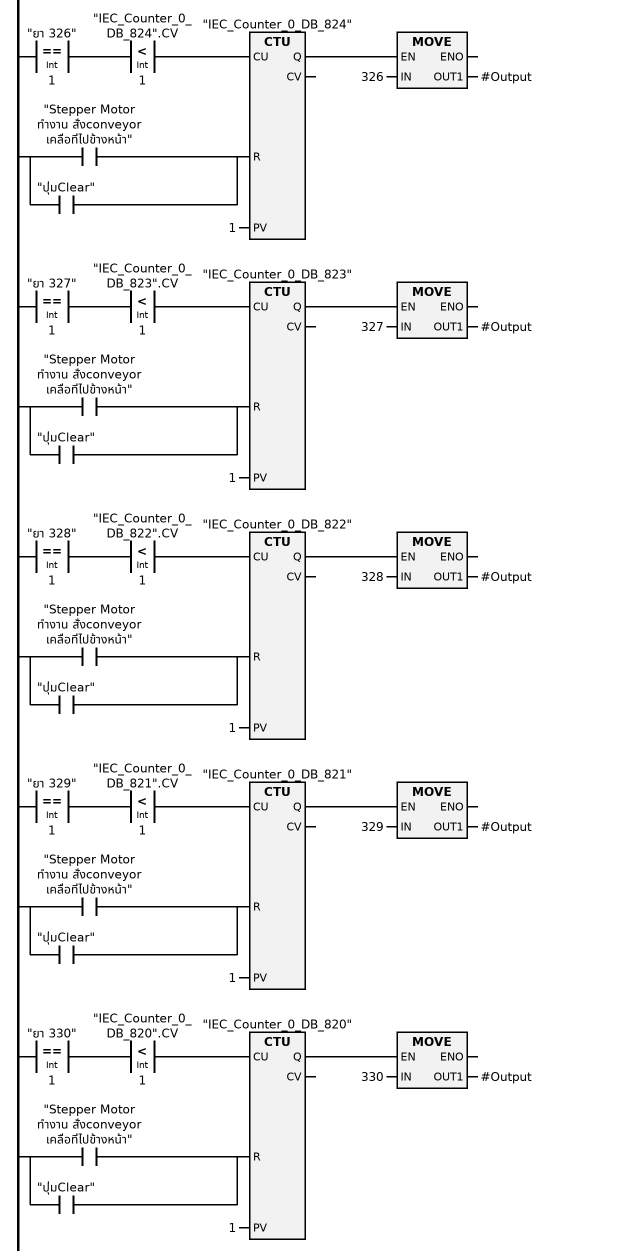
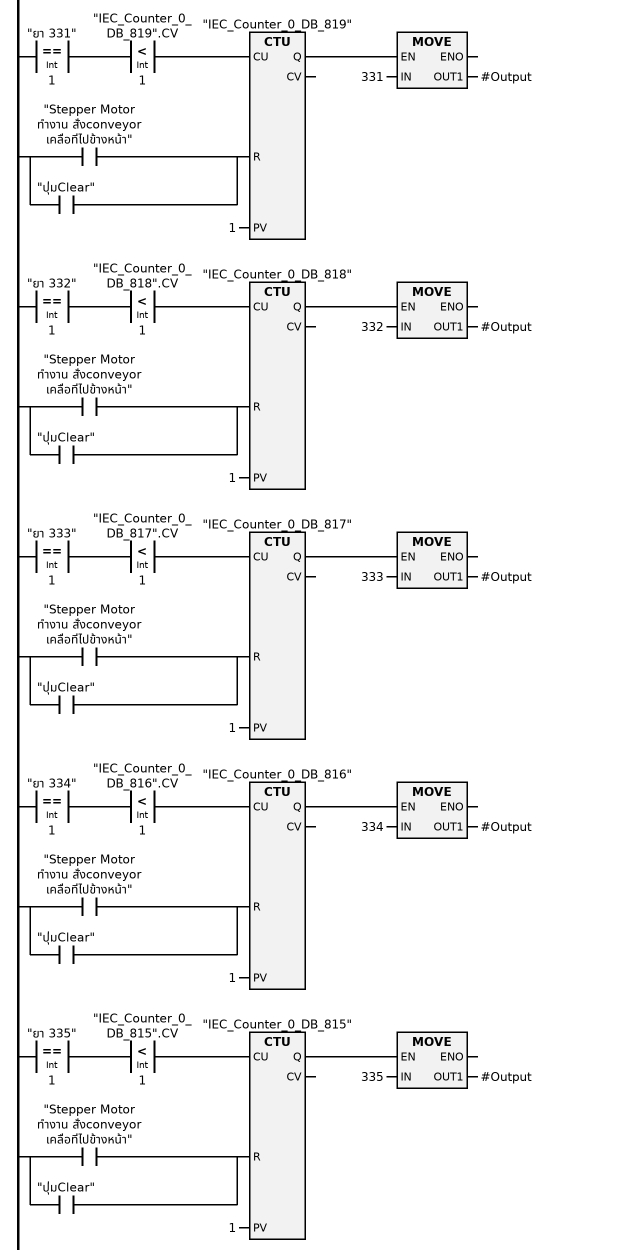
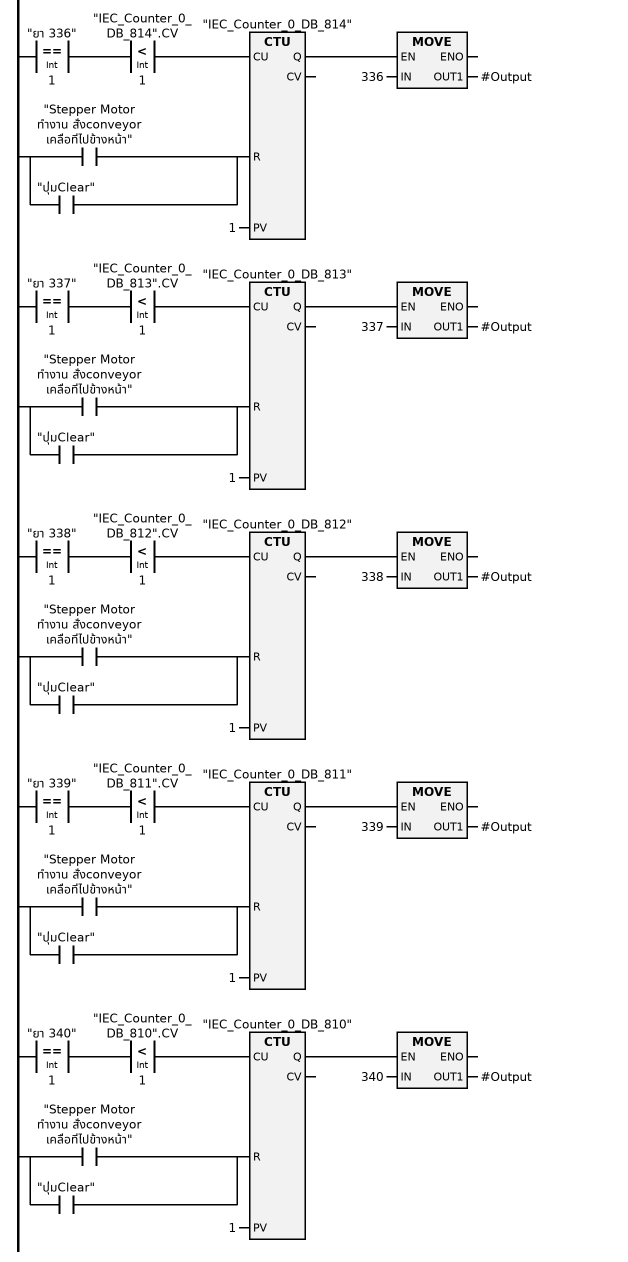
   "IEC_Counter_0_DB_829".CTU(CU := ("ยา 321" = 1) AND ("IEC_Counter_0_DB_829".CV < 1),
                           R := "Stepper Motor ทำงาน สั่งconveyor เคลื่อที่ไปข้างหน้า" OR "ปุ่มClear",
                           PV := 1);
   IF "IEC_Counter_0_DB_829".Q THEN #Output := 321; END_IF;
   "IEC_Counter_0_DB_828".CTU(CU := ("ยา 322" = 1) AND ("IEC_Counter_0_DB_828".CV < 1),
                           R := "Stepper Motor ทำงาน สั่งconveyor เคลื่อที่ไปข้างหน้า" OR "ปุ่มClear",
                           PV := 1);
   IF "IEC_Counter_0_DB_828".Q THEN #Output := 322; END_IF;
   "IEC_Counter_0_DB_825".CTU(CU := ("ยา 323" = 1) AND ("IEC_Counter_0_DB_825".CV < 1),
                           R := "Stepper Motor ทำงาน สั่งconveyor เคลื่อที่ไปข้างหน้า" OR "ปุ่มClear",
                           PV := 1);
   IF "IEC_Counter_0_DB_825".Q THEN #Output := 323; END_IF;
   "IEC_Counter_0_DB_827".CTU(CU := ("ยา 324" = 1) AND ("IEC_Counter_0_DB_827".CV < 1),
                           R := "Stepper Motor ทำงาน สั่งconveyor เคลื่อที่ไปข้างหน้า" OR "ปุ่มClear",
                           PV := 1);
   IF "IEC_Counter_0_DB_827".Q THEN #Output := 324; END_IF;
   "IEC_Counter_0_DB_826".CTU(CU := ("ยา 325" = 1) AND ("IEC_Counter_0_DB_826".CV < 1),
                           R := "Stepper Motor ทำงาน สั่งconveyor เคลื่อที่ไปข้างหน้า" OR "ปุ่มClear",
                           PV := 1);
   IF "IEC_Counter_0_DB_826".Q THEN #Output := 325; END_IF;
   "IEC_Counter_0_DB_824".CTU(CU := ("ยา 326" = 1) AND ("IEC_Counter_0_DB_824".CV < 1),
                           R := "Stepper Motor ทำงาน สั่งconveyor เคลื่อที่ไปข้างหน้า" OR "ปุ่มClear",
                           PV := 1);
   IF "IEC_Counter_0_DB_824".Q THEN #Output := 326; END_IF;
   "IEC_Counter_0_DB_823".CTU(CU := ("ยา 327" = 1) AND ("IEC_Counter_0_DB_823".CV < 1),
                           R := "Stepper Motor ทำงาน สั่งconveyor เคลื่อที่ไปข้างหน้า" OR "ปุ่มClear",
                           PV := 1);
   IF "IEC_Counter_0_DB_823".Q THEN #Output := 327; END_IF;
   "IEC_Counter_0_DB_822".CTU(CU := ("ยา 328" = 1) AND ("IEC_Counter_0_DB_822".CV < 1),
                           R := "Stepper Motor ทำงาน สั่งconveyor เคลื่อที่ไปข้างหน้า" OR "ปุ่มClear",
                           PV := 1);
   IF "IEC_Counter_0_DB_822".Q THEN #Output := 328; END_IF;
   "IEC_Counter_0_DB_821".CTU(CU := ("ยา 329" = 1) AND ("IEC_Counter_0_DB_821".CV < 1),
                           R := "Stepper Motor ทำงาน สั่งconveyor เคลื่อที่ไปข้างหน้า" OR "ปุ่มClear",
                           PV := 1);
   IF "IEC_Counter_0_DB_821".Q THEN #Output := 329; END_IF;
   "IEC_Counter_0_DB_820".CTU(CU := ("ยา 330" = 1) AND ("IEC_Counter_0_DB_820".CV < 1),
                           R := "Stepper Motor ทำงาน สั่งconveyor เคลื่อที่ไปข้างหน้า" OR "ปุ่มClear",
                           PV := 1);
   IF "IEC_Counter_0_DB_820".Q THEN #Output := 330; END_IF;
   "IEC_Counter_0_DB_819".CTU(CU := ("ยา 331" = 1) AND ("IEC_Counter_0_DB_819".CV < 1),
                           R := "Stepper Motor ทำงาน สั่งconveyor เคลื่อที่ไปข้างหน้า" OR "ปุ่มClear",
                           PV := 1);
   IF "IEC_Counter_0_DB_819".Q THEN #Output := 331; END_IF;
   "IEC_Counter_0_DB_818".CTU(CU := ("ยา 332" = 1) AND ("IEC_Counter_0_DB_818".CV < 1),
                           R := "Stepper Motor ทำงาน สั่งconveyor เคลื่อที่ไปข้างหน้า" OR "ปุ่มClear",
                           PV := 1);
   IF "IEC_Counter_0_DB_818".Q THEN #Output := 332; END_IF;
   "IEC_Counter_0_DB_817".CTU(CU := ("ยา 333" = 1) AND ("IEC_Counter_0_DB_817".CV < 1),
                           R := "Stepper Motor ทำงาน สั่งconveyor เคลื่อที่ไปข้างหน้า" OR "ปุ่มClear",
                           PV := 1);
   IF "IEC_Counter_0_DB_817".Q THEN #Output := 333; END_IF;
   "IEC_Counter_0_DB_816".CTU(CU := ("ยา 334" = 1) AND ("IEC_Counter_0_DB_816".CV < 1),
                           R := "Stepper Motor ทำงาน สั่งconveyor เคลื่อที่ไปข้างหน้า" OR "ปุ่มClear",
                           PV := 1);
   IF "IEC_Counter_0_DB_816".Q THEN #Output := 334; END_IF;
   "IEC_Counter_0_DB_815".CTU(CU := ("ยา 335" = 1) AND ("IEC_Counter_0_DB_815".CV < 1),
                           R := "Stepper Motor ทำงาน สั่งconveyor เคลื่อที่ไปข้างหน้า" OR "ปุ่มClear",
                           PV := 1);
   IF "IEC_Counter_0_DB_815".Q THEN #Output := 335; END_IF;
   "IEC_Counter_0_DB_814".CTU(CU := ("ยา 336" = 1) AND ("IEC_Counter_0_DB_814".CV < 1),
                           R := "Stepper Motor ทำงาน สั่งconveyor เคลื่อที่ไปข้างหน้า" OR "ปุ่มClear",
                           PV := 1);
   IF "IEC_Counter_0_DB_814".Q THEN #Output := 336; END_IF;
   "IEC_Counter_0_DB_813".CTU(CU := ("ยา 337" = 1) AND ("IEC_Counter_0_DB_813".CV < 1),
                           R := "Stepper Motor ทำงาน สั่งconveyor เคลื่อที่ไปข้างหน้า" OR "ปุ่มClear",
                           PV := 1);
   IF "IEC_Counter_0_DB_813".Q THEN #Output := 337; END_IF;
   "IEC_Counter_0_DB_812".CTU(CU := ("ยา 338" = 1) AND ("IEC_Counter_0_DB_812".CV < 1),
                           R := "Stepper Motor ทำงาน สั่งconveyor เคลื่อที่ไปข้างหน้า" OR "ปุ่มClear",
                           PV := 1);
   IF "IEC_Counter_0_DB_812".Q THEN #Output := 338; END_IF;
   "IEC_Counter_0_DB_811".CTU(CU := ("ยา 339" = 1) AND ("IEC_Counter_0_DB_811".CV < 1),
                           R := "Stepper Motor ทำงาน สั่งconveyor เคลื่อที่ไปข้างหน้า" OR "ปุ่มClear",
                           PV := 1);
   IF "IEC_Counter_0_DB_811".Q THEN #Output := 339; END_IF;
   "IEC_Counter_0_DB_810".CTU(CU := ("ยา 340" = 1) AND ("IEC_Counter_0_DB_810".CV < 1),
                           R := "Stepper Motor ทำงาน สั่งconveyor เคลื่อที่ไปข้างหน้า" OR "ปุ่มClear",
                           PV := 1);
   IF "IEC_Counter_0_DB_810".Q THEN #Output := 340; END_IF;
END_REGION

REGION Network 18
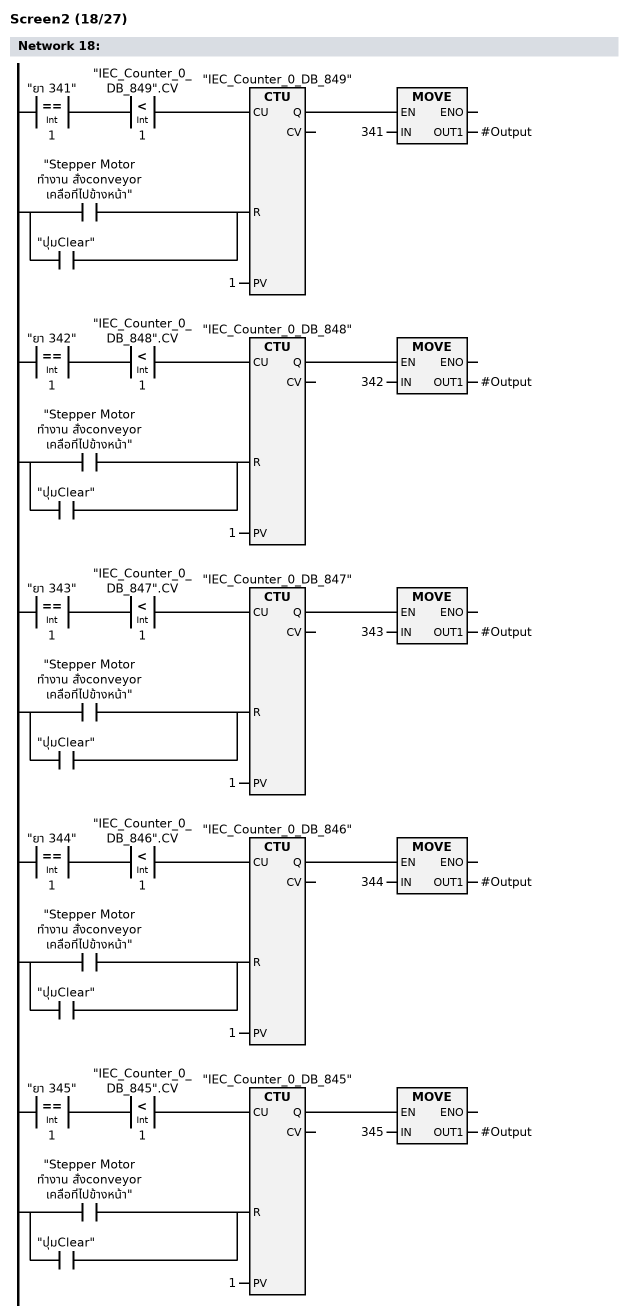
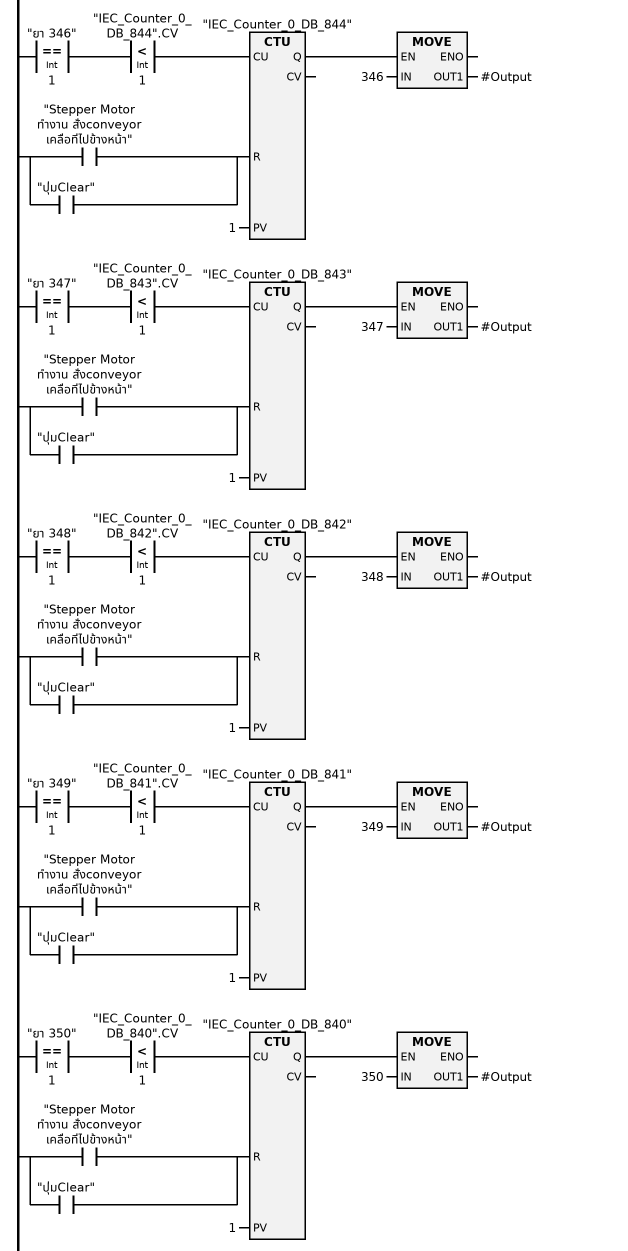
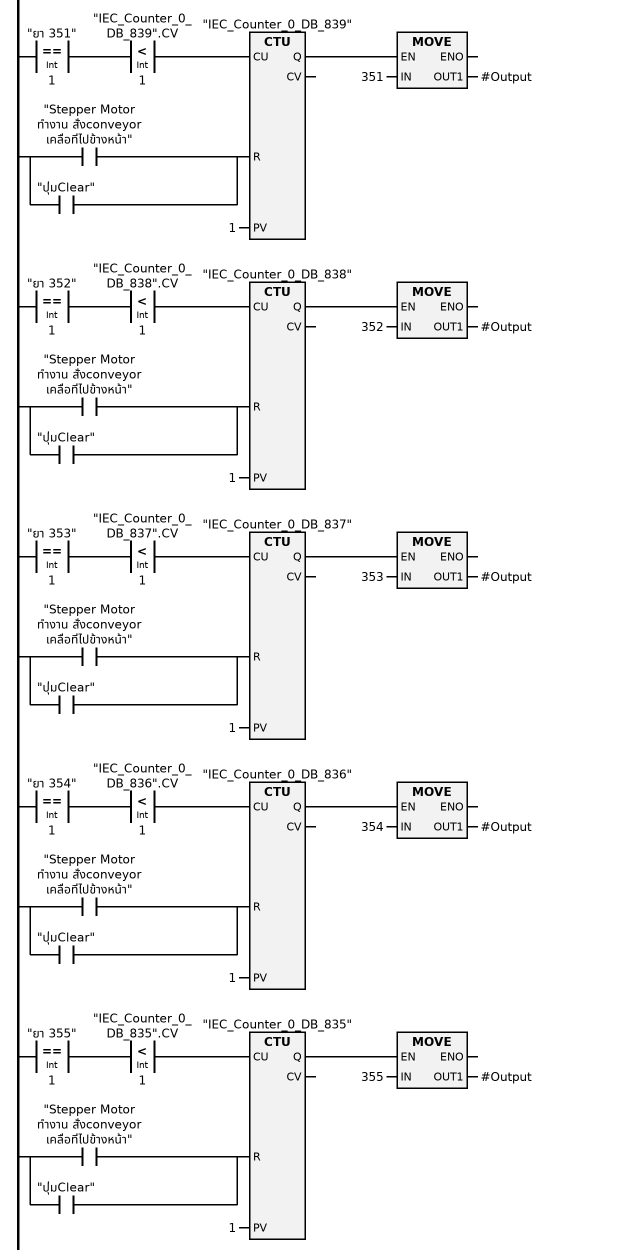
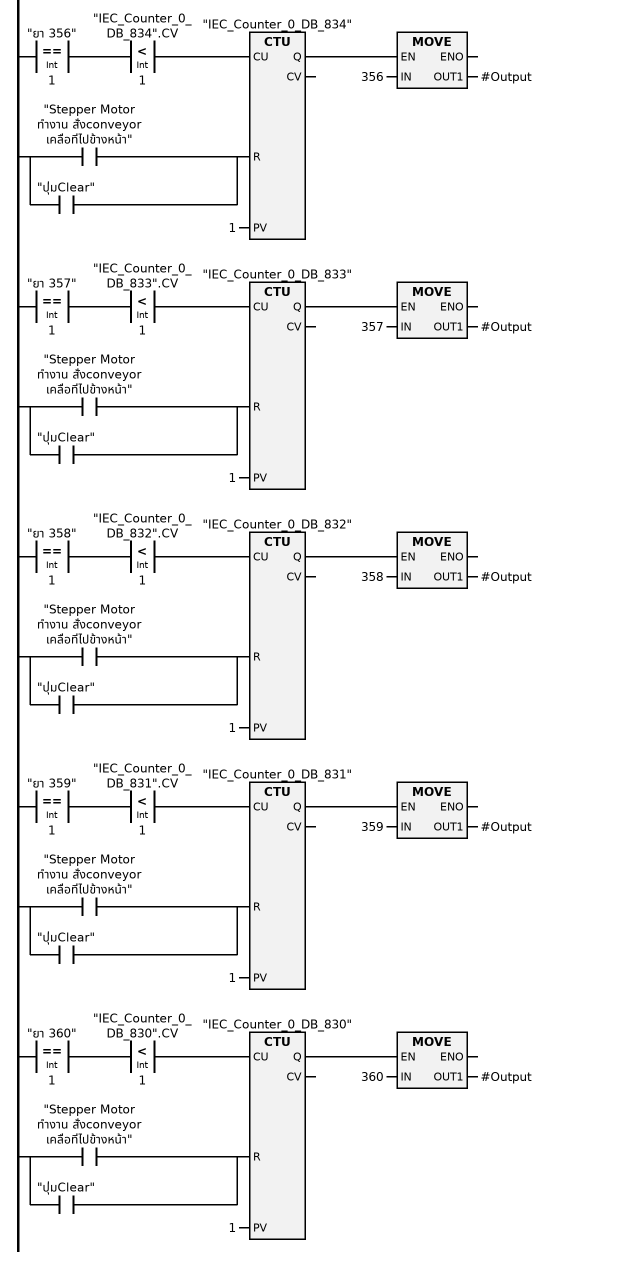
   "IEC_Counter_0_DB_849".CTU(CU := ("ยา 341" = 1) AND ("IEC_Counter_0_DB_849".CV < 1),
                           R := "Stepper Motor ทำงาน สั่งconveyor เคลื่อที่ไปข้างหน้า" OR "ปุ่มClear",
                           PV := 1);
   IF "IEC_Counter_0_DB_849".Q THEN #Output := 341; END_IF;
   "IEC_Counter_0_DB_848".CTU(CU := ("ยา 342" = 1) AND ("IEC_Counter_0_DB_848".CV < 1),
                           R := "Stepper Motor ทำงาน สั่งconveyor เคลื่อที่ไปข้างหน้า" OR "ปุ่มClear",
                           PV := 1);
   IF "IEC_Counter_0_DB_848".Q THEN #Output := 342; END_IF;
   "IEC_Counter_0_DB_847".CTU(CU := ("ยา 343" = 1) AND ("IEC_Counter_0_DB_847".CV < 1),
                           R := "Stepper Motor ทำงาน สั่งconveyor เคลื่อที่ไปข้างหน้า" OR "ปุ่มClear",
                           PV := 1);
   IF "IEC_Counter_0_DB_847".Q THEN #Output := 343; END_IF;
   "IEC_Counter_0_DB_846".CTU(CU := ("ยา 344" = 1) AND ("IEC_Counter_0_DB_846".CV < 1),
                           R := "Stepper Motor ทำงาน สั่งconveyor เคลื่อที่ไปข้างหน้า" OR "ปุ่มClear",
                           PV := 1);
   IF "IEC_Counter_0_DB_846".Q THEN #Output := 344; END_IF;
   "IEC_Counter_0_DB_845".CTU(CU := ("ยา 345" = 1) AND ("IEC_Counter_0_DB_845".CV < 1),
                           R := "Stepper Motor ทำงาน สั่งconveyor เคลื่อที่ไปข้างหน้า" OR "ปุ่มClear",
                           PV := 1);
   IF "IEC_Counter_0_DB_845".Q THEN #Output := 345; END_IF;
   "IEC_Counter_0_DB_844".CTU(CU := ("ยา 346" = 1) AND ("IEC_Counter_0_DB_844".CV < 1),
                           R := "Stepper Motor ทำงาน สั่งconveyor เคลื่อที่ไปข้างหน้า" OR "ปุ่มClear",
                           PV := 1);
   IF "IEC_Counter_0_DB_844".Q THEN #Output := 346; END_IF;
   "IEC_Counter_0_DB_843".CTU(CU := ("ยา 347" = 1) AND ("IEC_Counter_0_DB_843".CV < 1),
                           R := "Stepper Motor ทำงาน สั่งconveyor เคลื่อที่ไปข้างหน้า" OR "ปุ่มClear",
                           PV := 1);
   IF "IEC_Counter_0_DB_843".Q THEN #Output := 347; END_IF;
   "IEC_Counter_0_DB_842".CTU(CU := ("ยา 348" = 1) AND ("IEC_Counter_0_DB_842".CV < 1),
                           R := "Stepper Motor ทำงาน สั่งconveyor เคลื่อที่ไปข้างหน้า" OR "ปุ่มClear",
                           PV := 1);
   IF "IEC_Counter_0_DB_842".Q THEN #Output := 348; END_IF;
   "IEC_Counter_0_DB_841".CTU(CU := ("ยา 349" = 1) AND ("IEC_Counter_0_DB_841".CV < 1),
                           R := "Stepper Motor ทำงาน สั่งconveyor เคลื่อที่ไปข้างหน้า" OR "ปุ่มClear",
                           PV := 1);
   IF "IEC_Counter_0_DB_841".Q THEN #Output := 349; END_IF;
   "IEC_Counter_0_DB_840".CTU(CU := ("ยา 350" = 1) AND ("IEC_Counter_0_DB_840".CV < 1),
                           R := "Stepper Motor ทำงาน สั่งconveyor เคลื่อที่ไปข้างหน้า" OR "ปุ่มClear",
                           PV := 1);
   IF "IEC_Counter_0_DB_840".Q THEN #Output := 350; END_IF;
   "IEC_Counter_0_DB_839".CTU(CU := ("ยา 351" = 1) AND ("IEC_Counter_0_DB_839".CV < 1),
                           R := "Stepper Motor ทำงาน สั่งconveyor เคลื่อที่ไปข้างหน้า" OR "ปุ่มClear",
                           PV := 1);
   IF "IEC_Counter_0_DB_839".Q THEN #Output := 351; END_IF;
   "IEC_Counter_0_DB_838".CTU(CU := ("ยา 352" = 1) AND ("IEC_Counter_0_DB_838".CV < 1),
                           R := "Stepper Motor ทำงาน สั่งconveyor เคลื่อที่ไปข้างหน้า" OR "ปุ่มClear",
                           PV := 1);
   IF "IEC_Counter_0_DB_838".Q THEN #Output := 352; END_IF;
   "IEC_Counter_0_DB_837".CTU(CU := ("ยา 353" = 1) AND ("IEC_Counter_0_DB_837".CV < 1),
                           R := "Stepper Motor ทำงาน สั่งconveyor เคลื่อที่ไปข้างหน้า" OR "ปุ่มClear",
                           PV := 1);
   IF "IEC_Counter_0_DB_837".Q THEN #Output := 353; END_IF;
   "IEC_Counter_0_DB_836".CTU(CU := ("ยา 354" = 1) AND ("IEC_Counter_0_DB_836".CV < 1),
                           R := "Stepper Motor ทำงาน สั่งconveyor เคลื่อที่ไปข้างหน้า" OR "ปุ่มClear",
                           PV := 1);
   IF "IEC_Counter_0_DB_836".Q THEN #Output := 354; END_IF;
   "IEC_Counter_0_DB_835".CTU(CU := ("ยา 355" = 1) AND ("IEC_Counter_0_DB_835".CV < 1),
                           R := "Stepper Motor ทำงาน สั่งconveyor เคลื่อที่ไปข้างหน้า" OR "ปุ่มClear",
                           PV := 1);
   IF "IEC_Counter_0_DB_835".Q THEN #Output := 355; END_IF;
   "IEC_Counter_0_DB_834".CTU(CU := ("ยา 356" = 1) AND ("IEC_Counter_0_DB_834".CV < 1),
                           R := "Stepper Motor ทำงาน สั่งconveyor เคลื่อที่ไปข้างหน้า" OR "ปุ่มClear",
                           PV := 1);
   IF "IEC_Counter_0_DB_834".Q THEN #Output := 356; END_IF;
   "IEC_Counter_0_DB_833".CTU(CU := ("ยา 357" = 1) AND ("IEC_Counter_0_DB_833".CV < 1),
                           R := "Stepper Motor ทำงาน สั่งconveyor เคลื่อที่ไปข้างหน้า" OR "ปุ่มClear",
                           PV := 1);
   IF "IEC_Counter_0_DB_833".Q THEN #Output := 357; END_IF;
   "IEC_Counter_0_DB_832".CTU(CU := ("ยา 358" = 1) AND ("IEC_Counter_0_DB_832".CV < 1),
                           R := "Stepper Motor ทำงาน สั่งconveyor เคลื่อที่ไปข้างหน้า" OR "ปุ่มClear",
                           PV := 1);
   IF "IEC_Counter_0_DB_832".Q THEN #Output := 358; END_IF;
   "IEC_Counter_0_DB_831".CTU(CU := ("ยา 359" = 1) AND ("IEC_Counter_0_DB_831".CV < 1),
                           R := "Stepper Motor ทำงาน สั่งconveyor เคลื่อที่ไปข้างหน้า" OR "ปุ่มClear",
                           PV := 1);
   IF "IEC_Counter_0_DB_831".Q THEN #Output := 359; END_IF;
   "IEC_Counter_0_DB_830".CTU(CU := ("ยา 360" = 1) AND ("IEC_Counter_0_DB_830".CV < 1),
                           R := "Stepper Motor ทำงาน สั่งconveyor เคลื่อที่ไปข้างหน้า" OR "ปุ่มClear",
                           PV := 1);
   IF "IEC_Counter_0_DB_830".Q THEN #Output := 360; END_IF;
END_REGION

REGION Network 19
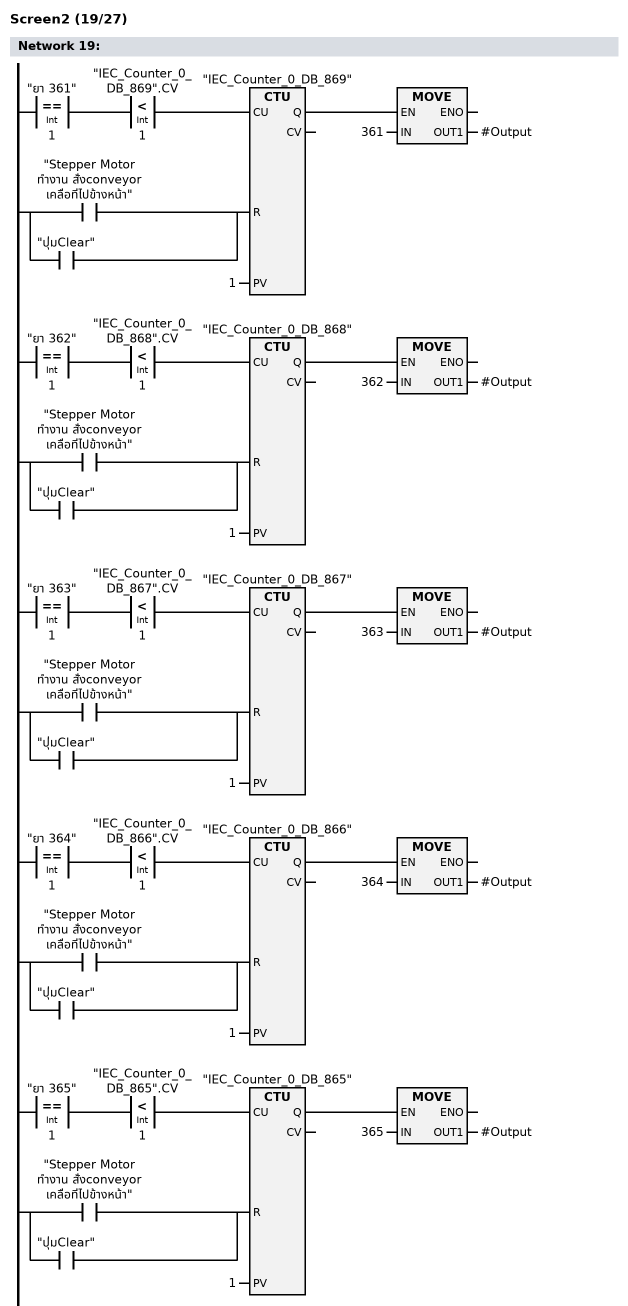
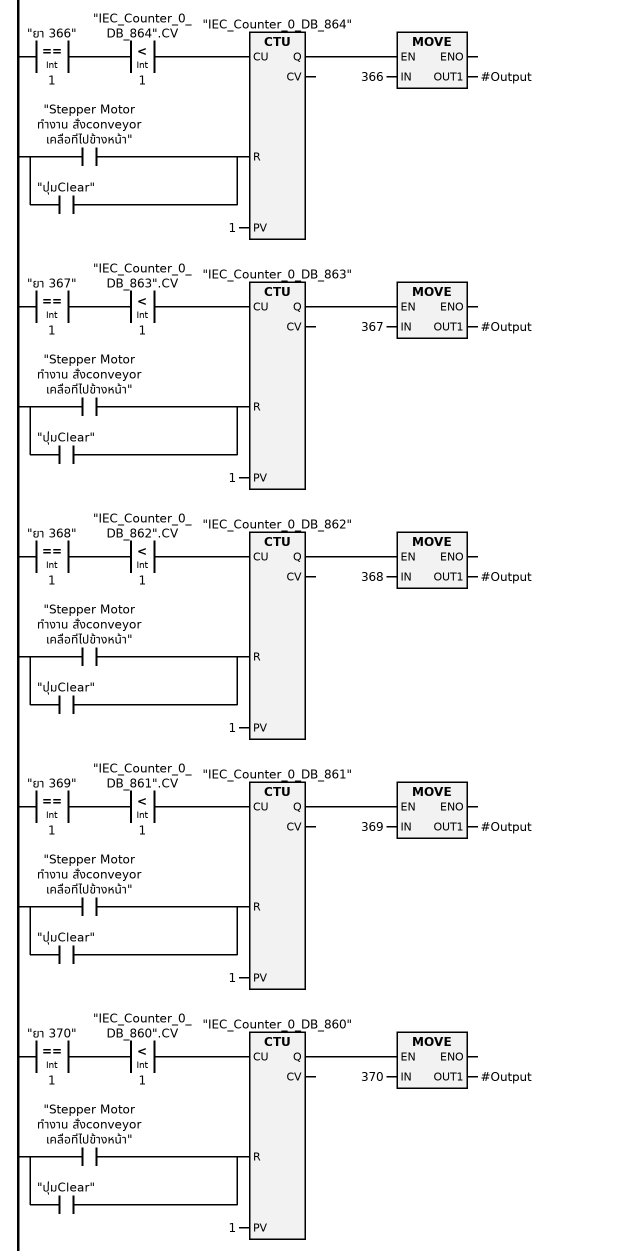
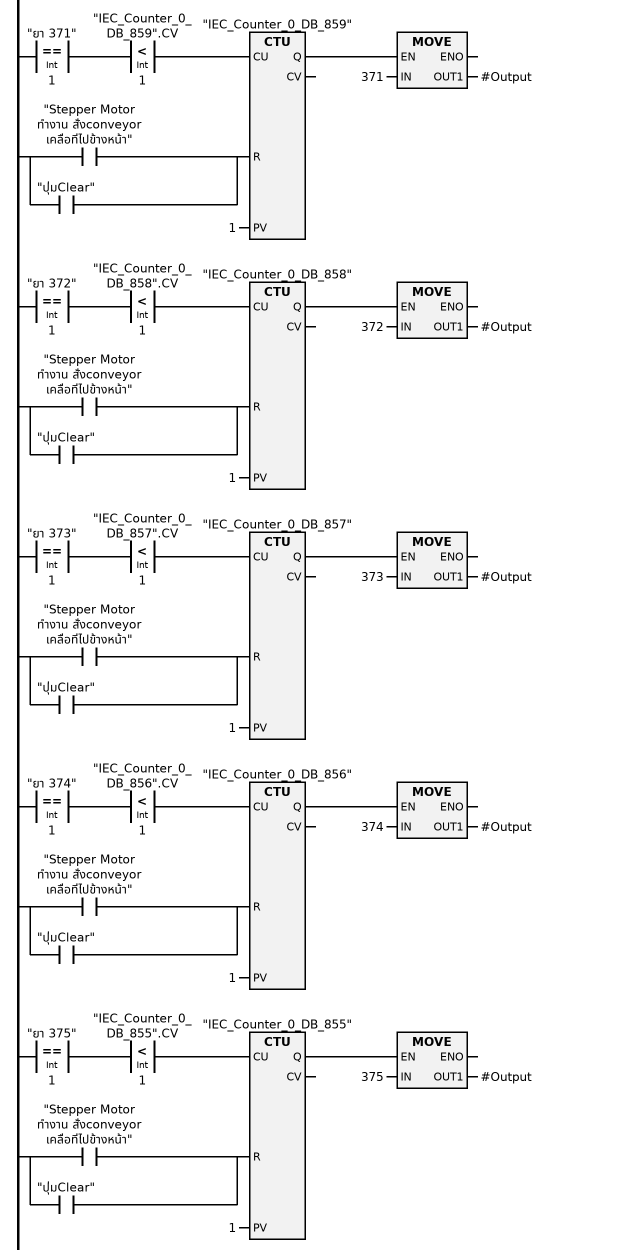
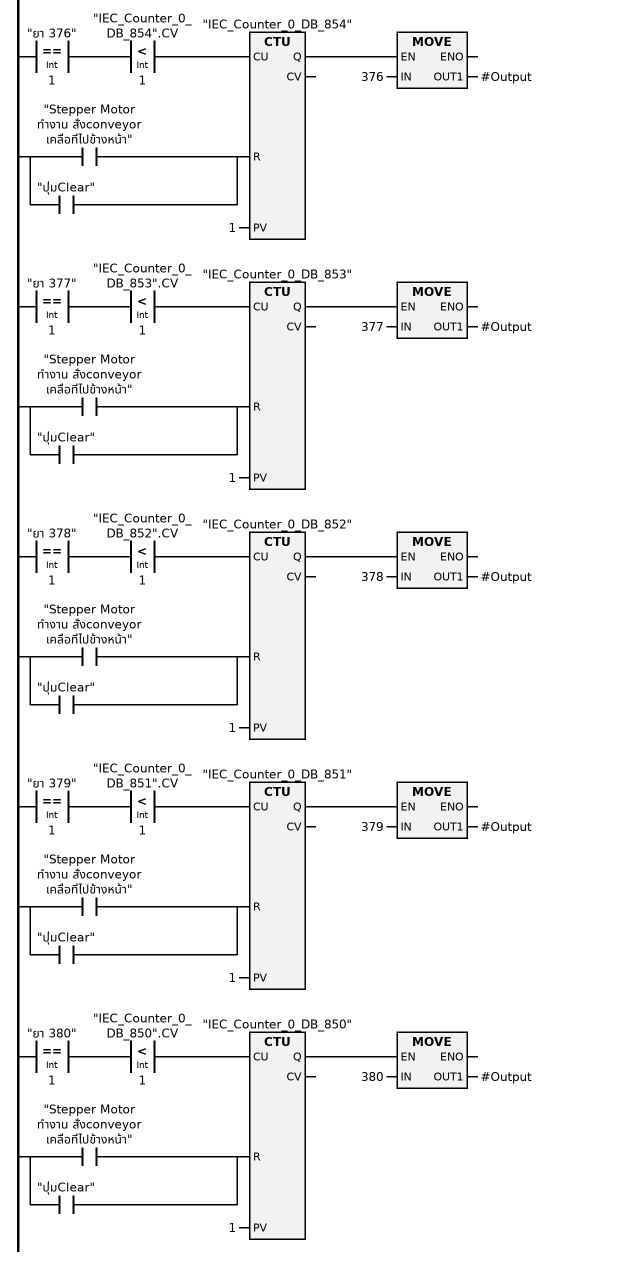
   "IEC_Counter_0_DB_869".CTU(CU := ("ยา 361" = 1) AND ("IEC_Counter_0_DB_869".CV < 1),
                           R := "Stepper Motor ทำงาน สั่งconveyor เคลื่อที่ไปข้างหน้า" OR "ปุ่มClear",
                           PV := 1);
   IF "IEC_Counter_0_DB_869".Q THEN #Output := 361; END_IF;
   "IEC_Counter_0_DB_868".CTU(CU := ("ยา 362" = 1) AND ("IEC_Counter_0_DB_868".CV < 1),
                           R := "Stepper Motor ทำงาน สั่งconveyor เคลื่อที่ไปข้างหน้า" OR "ปุ่มClear",
                           PV := 1);
   IF "IEC_Counter_0_DB_868".Q THEN #Output := 362; END_IF;
   "IEC_Counter_0_DB_867".CTU(CU := ("ยา 363" = 1) AND ("IEC_Counter_0_DB_867".CV < 1),
                           R := "Stepper Motor ทำงาน สั่งconveyor เคลื่อที่ไปข้างหน้า" OR "ปุ่มClear",
                           PV := 1);
   IF "IEC_Counter_0_DB_867".Q THEN #Output := 363; END_IF;
   "IEC_Counter_0_DB_866".CTU(CU := ("ยา 364" = 1) AND ("IEC_Counter_0_DB_866".CV < 1),
                           R := "Stepper Motor ทำงาน สั่งconveyor เคลื่อที่ไปข้างหน้า" OR "ปุ่มClear",
                           PV := 1);
   IF "IEC_Counter_0_DB_866".Q THEN #Output := 364; END_IF;
   "IEC_Counter_0_DB_865".CTU(CU := ("ยา 365" = 1) AND ("IEC_Counter_0_DB_865".CV < 1),
                           R := "Stepper Motor ทำงาน สั่งconveyor เคลื่อที่ไปข้างหน้า" OR "ปุ่มClear",
                           PV := 1);
   IF "IEC_Counter_0_DB_865".Q THEN #Output := 365; END_IF;
   "IEC_Counter_0_DB_864".CTU(CU := ("ยา 366" = 1) AND ("IEC_Counter_0_DB_864".CV < 1),
                           R := "Stepper Motor ทำงาน สั่งconveyor เคลื่อที่ไปข้างหน้า" OR "ปุ่มClear",
                           PV := 1);
   IF "IEC_Counter_0_DB_864".Q THEN #Output := 366; END_IF;
   "IEC_Counter_0_DB_863".CTU(CU := ("ยา 367" = 1) AND ("IEC_Counter_0_DB_863".CV < 1),
                           R := "Stepper Motor ทำงาน สั่งconveyor เคลื่อที่ไปข้างหน้า" OR "ปุ่มClear",
                           PV := 1);
   IF "IEC_Counter_0_DB_863".Q THEN #Output := 367; END_IF;
   "IEC_Counter_0_DB_862".CTU(CU := ("ยา 368" = 1) AND ("IEC_Counter_0_DB_862".CV < 1),
                           R := "Stepper Motor ทำงาน สั่งconveyor เคลื่อที่ไปข้างหน้า" OR "ปุ่มClear",
                           PV := 1);
   IF "IEC_Counter_0_DB_862".Q THEN #Output := 368; END_IF;
   "IEC_Counter_0_DB_861".CTU(CU := ("ยา 369" = 1) AND ("IEC_Counter_0_DB_861".CV < 1),
                           R := "Stepper Motor ทำงาน สั่งconveyor เคลื่อที่ไปข้างหน้า" OR "ปุ่มClear",
                           PV := 1);
   IF "IEC_Counter_0_DB_861".Q THEN #Output := 369; END_IF;
   "IEC_Counter_0_DB_860".CTU(CU := ("ยา 370" = 1) AND ("IEC_Counter_0_DB_860".CV < 1),
                           R := "Stepper Motor ทำงาน สั่งconveyor เคลื่อที่ไปข้างหน้า" OR "ปุ่มClear",
                           PV := 1);
   IF "IEC_Counter_0_DB_860".Q THEN #Output := 370; END_IF;
   "IEC_Counter_0_DB_859".CTU(CU := ("ยา 371" = 1) AND ("IEC_Counter_0_DB_859".CV < 1),
                           R := "Stepper Motor ทำงาน สั่งconveyor เคลื่อที่ไปข้างหน้า" OR "ปุ่มClear",
                           PV := 1);
   IF "IEC_Counter_0_DB_859".Q THEN #Output := 371; END_IF;
   "IEC_Counter_0_DB_858".CTU(CU := ("ยา 372" = 1) AND ("IEC_Counter_0_DB_858".CV < 1),
                           R := "Stepper Motor ทำงาน สั่งconveyor เคลื่อที่ไปข้างหน้า" OR "ปุ่มClear",
                           PV := 1);
   IF "IEC_Counter_0_DB_858".Q THEN #Output := 372; END_IF;
   "IEC_Counter_0_DB_857".CTU(CU := ("ยา 373" = 1) AND ("IEC_Counter_0_DB_857".CV < 1),
                           R := "Stepper Motor ทำงาน สั่งconveyor เคลื่อที่ไปข้างหน้า" OR "ปุ่มClear",
                           PV := 1);
   IF "IEC_Counter_0_DB_857".Q THEN #Output := 373; END_IF;
   "IEC_Counter_0_DB_856".CTU(CU := ("ยา 374" = 1) AND ("IEC_Counter_0_DB_856".CV < 1),
                           R := "Stepper Motor ทำงาน สั่งconveyor เคลื่อที่ไปข้างหน้า" OR "ปุ่มClear",
                           PV := 1);
   IF "IEC_Counter_0_DB_856".Q THEN #Output := 374; END_IF;
   "IEC_Counter_0_DB_855".CTU(CU := ("ยา 375" = 1) AND ("IEC_Counter_0_DB_855".CV < 1),
                           R := "Stepper Motor ทำงาน สั่งconveyor เคลื่อที่ไปข้างหน้า" OR "ปุ่มClear",
                           PV := 1);
   IF "IEC_Counter_0_DB_855".Q THEN #Output := 375; END_IF;
   "IEC_Counter_0_DB_854".CTU(CU := ("ยา 376" = 1) AND ("IEC_Counter_0_DB_854".CV < 1),
                           R := "Stepper Motor ทำงาน สั่งconveyor เคลื่อที่ไปข้างหน้า" OR "ปุ่มClear",
                           PV := 1);
   IF "IEC_Counter_0_DB_854".Q THEN #Output := 376; END_IF;
   "IEC_Counter_0_DB_853".CTU(CU := ("ยา 377" = 1) AND ("IEC_Counter_0_DB_853".CV < 1),
                           R := "Stepper Motor ทำงาน สั่งconveyor เคลื่อที่ไปข้างหน้า" OR "ปุ่มClear",
                           PV := 1);
   IF "IEC_Counter_0_DB_853".Q THEN #Output := 377; END_IF;
   "IEC_Counter_0_DB_852".CTU(CU := ("ยา 378" = 1) AND ("IEC_Counter_0_DB_852".CV < 1),
                           R := "Stepper Motor ทำงาน สั่งconveyor เคลื่อที่ไปข้างหน้า" OR "ปุ่มClear",
                           PV := 1);
   IF "IEC_Counter_0_DB_852".Q THEN #Output := 378; END_IF;
   "IEC_Counter_0_DB_851".CTU(CU := ("ยา 379" = 1) AND ("IEC_Counter_0_DB_851".CV < 1),
                           R := "Stepper Motor ทำงาน สั่งconveyor เคลื่อที่ไปข้างหน้า" OR "ปุ่มClear",
                           PV := 1);
   IF "IEC_Counter_0_DB_851".Q THEN #Output := 379; END_IF;
   "IEC_Counter_0_DB_850".CTU(CU := ("ยา 380" = 1) AND ("IEC_Counter_0_DB_850".CV < 1),
                           R := "Stepper Motor ทำงาน สั่งconveyor เคลื่อที่ไปข้างหน้า" OR "ปุ่มClear",
                           PV := 1);
   IF "IEC_Counter_0_DB_850".Q THEN #Output := 380; END_IF;
END_REGION

REGION Network 20
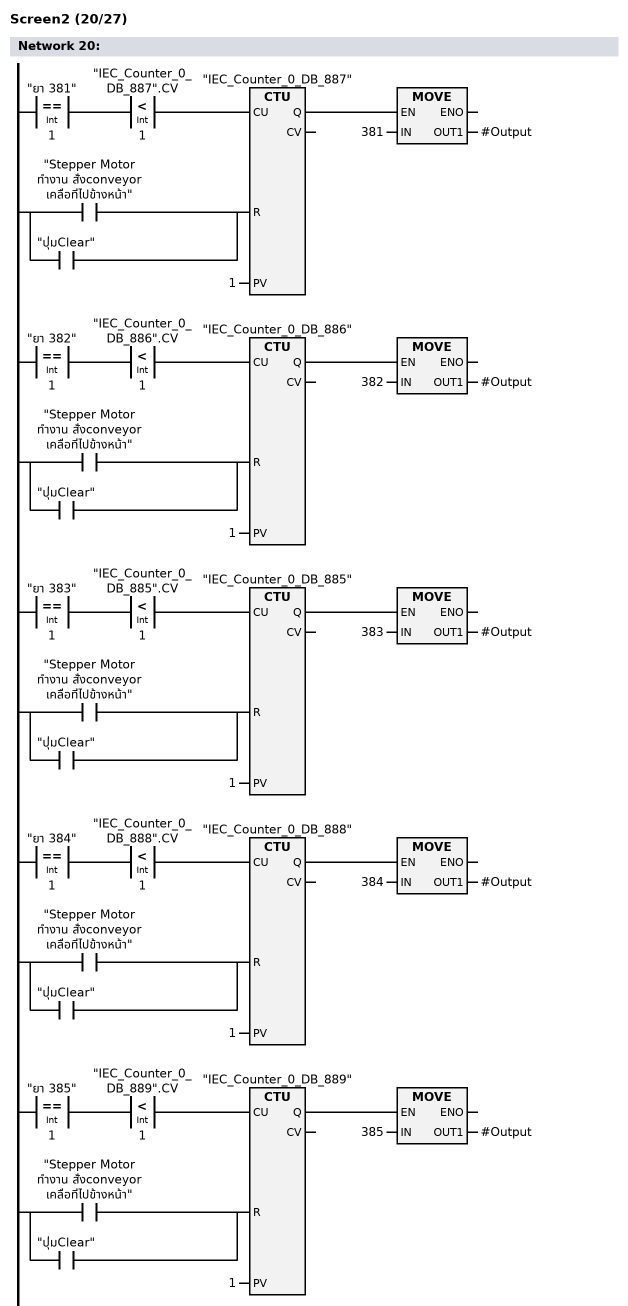
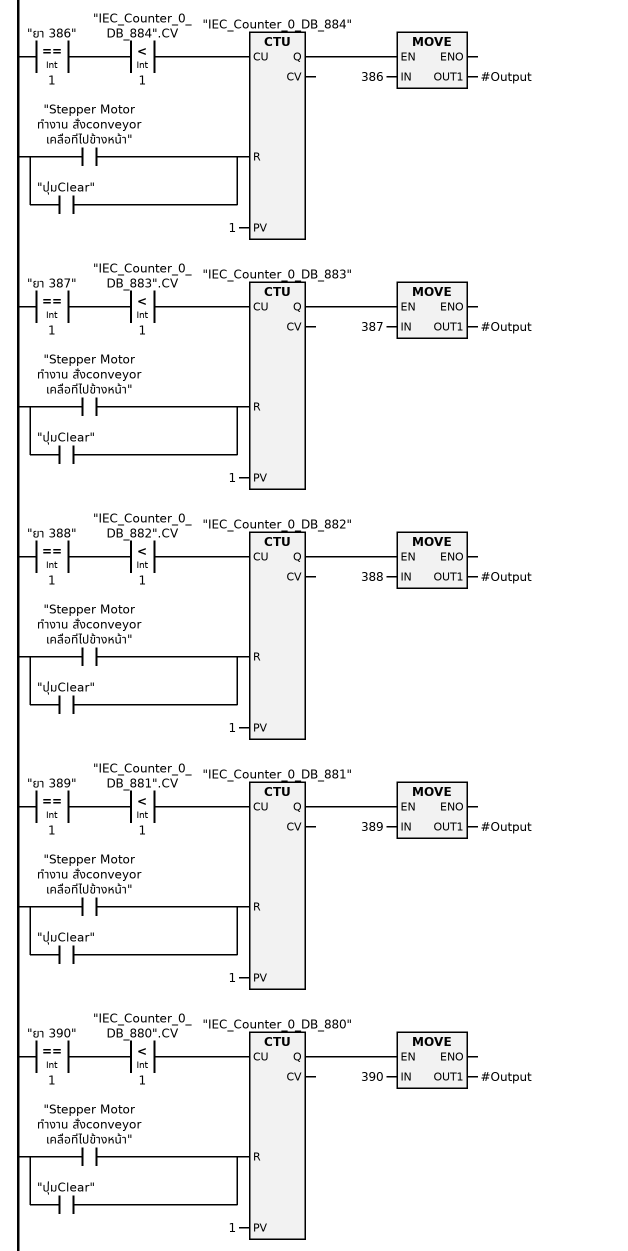
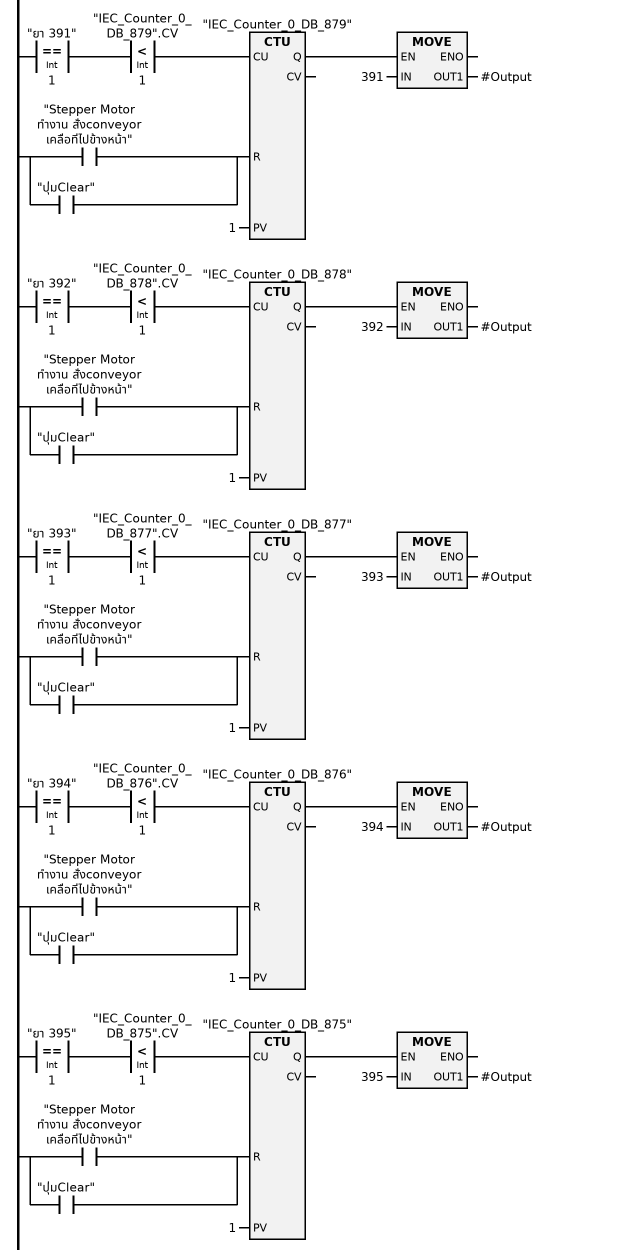
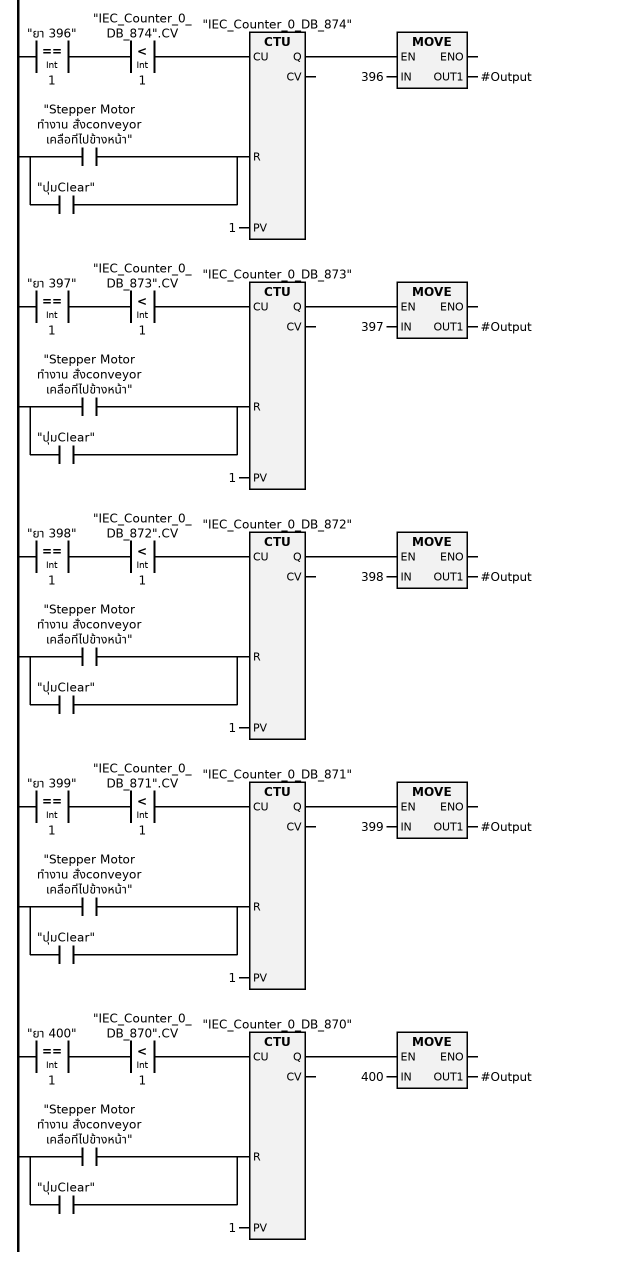
   "IEC_Counter_0_DB_887".CTU(CU := ("ยา 381" = 1) AND ("IEC_Counter_0_DB_887".CV < 1),
                           R := "Stepper Motor ทำงาน สั่งconveyor เคลื่อที่ไปข้างหน้า" OR "ปุ่มClear",
                           PV := 1);
   IF "IEC_Counter_0_DB_887".Q THEN #Output := 381; END_IF;
   "IEC_Counter_0_DB_886".CTU(CU := ("ยา 382" = 1) AND ("IEC_Counter_0_DB_886".CV < 1),
                           R := "Stepper Motor ทำงาน สั่งconveyor เคลื่อที่ไปข้างหน้า" OR "ปุ่มClear",
                           PV := 1);
   IF "IEC_Counter_0_DB_886".Q THEN #Output := 382; END_IF;
   "IEC_Counter_0_DB_885".CTU(CU := ("ยา 383" = 1) AND ("IEC_Counter_0_DB_885".CV < 1),
                           R := "Stepper Motor ทำงาน สั่งconveyor เคลื่อที่ไปข้างหน้า" OR "ปุ่มClear",
                           PV := 1);
   IF "IEC_Counter_0_DB_885".Q THEN #Output := 383; END_IF;
   "IEC_Counter_0_DB_888".CTU(CU := ("ยา 384" = 1) AND ("IEC_Counter_0_DB_888".CV < 1),
                           R := "Stepper Motor ทำงาน สั่งconveyor เคลื่อที่ไปข้างหน้า" OR "ปุ่มClear",
                           PV := 1);
   IF "IEC_Counter_0_DB_888".Q THEN #Output := 384; END_IF;
   "IEC_Counter_0_DB_889".CTU(CU := ("ยา 385" = 1) AND ("IEC_Counter_0_DB_889".CV < 1),
                           R := "Stepper Motor ทำงาน สั่งconveyor เคลื่อที่ไปข้างหน้า" OR "ปุ่มClear",
                           PV := 1);
   IF "IEC_Counter_0_DB_889".Q THEN #Output := 385; END_IF;
   "IEC_Counter_0_DB_884".CTU(CU := ("ยา 386" = 1) AND ("IEC_Counter_0_DB_884".CV < 1),
                           R := "Stepper Motor ทำงาน สั่งconveyor เคลื่อที่ไปข้างหน้า" OR "ปุ่มClear",
                           PV := 1);
   IF "IEC_Counter_0_DB_884".Q THEN #Output := 386; END_IF;
   "IEC_Counter_0_DB_883".CTU(CU := ("ยา 387" = 1) AND ("IEC_Counter_0_DB_883".CV < 1),
                           R := "Stepper Motor ทำงาน สั่งconveyor เคลื่อที่ไปข้างหน้า" OR "ปุ่มClear",
                           PV := 1);
   IF "IEC_Counter_0_DB_883".Q THEN #Output := 387; END_IF;
   "IEC_Counter_0_DB_882".CTU(CU := ("ยา 388" = 1) AND ("IEC_Counter_0_DB_882".CV < 1),
                           R := "Stepper Motor ทำงาน สั่งconveyor เคลื่อที่ไปข้างหน้า" OR "ปุ่มClear",
                           PV := 1);
   IF "IEC_Counter_0_DB_882".Q THEN #Output := 388; END_IF;
   "IEC_Counter_0_DB_881".CTU(CU := ("ยา 389" = 1) AND ("IEC_Counter_0_DB_881".CV < 1),
                           R := "Stepper Motor ทำงาน สั่งconveyor เคลื่อที่ไปข้างหน้า" OR "ปุ่มClear",
                           PV := 1);
   IF "IEC_Counter_0_DB_881".Q THEN #Output := 389; END_IF;
   "IEC_Counter_0_DB_880".CTU(CU := ("ยา 390" = 1) AND ("IEC_Counter_0_DB_880".CV < 1),
                           R := "Stepper Motor ทำงาน สั่งconveyor เคลื่อที่ไปข้างหน้า" OR "ปุ่มClear",
                           PV := 1);
   IF "IEC_Counter_0_DB_880".Q THEN #Output := 390; END_IF;
   "IEC_Counter_0_DB_879".CTU(CU := ("ยา 391" = 1) AND ("IEC_Counter_0_DB_879".CV < 1),
                           R := "Stepper Motor ทำงาน สั่งconveyor เคลื่อที่ไปข้างหน้า" OR "ปุ่มClear",
                           PV := 1);
   IF "IEC_Counter_0_DB_879".Q THEN #Output := 391; END_IF;
   "IEC_Counter_0_DB_878".CTU(CU := ("ยา 392" = 1) AND ("IEC_Counter_0_DB_878".CV < 1),
                           R := "Stepper Motor ทำงาน สั่งconveyor เคลื่อที่ไปข้างหน้า" OR "ปุ่มClear",
                           PV := 1);
   IF "IEC_Counter_0_DB_878".Q THEN #Output := 392; END_IF;
   "IEC_Counter_0_DB_877".CTU(CU := ("ยา 393" = 1) AND ("IEC_Counter_0_DB_877".CV < 1),
                           R := "Stepper Motor ทำงาน สั่งconveyor เคลื่อที่ไปข้างหน้า" OR "ปุ่มClear",
                           PV := 1);
   IF "IEC_Counter_0_DB_877".Q THEN #Output := 393; END_IF;
   "IEC_Counter_0_DB_876".CTU(CU := ("ยา 394" = 1) AND ("IEC_Counter_0_DB_876".CV < 1),
                           R := "Stepper Motor ทำงาน สั่งconveyor เคลื่อที่ไปข้างหน้า" OR "ปุ่มClear",
                           PV := 1);
   IF "IEC_Counter_0_DB_876".Q THEN #Output := 394; END_IF;
   "IEC_Counter_0_DB_875".CTU(CU := ("ยา 395" = 1) AND ("IEC_Counter_0_DB_875".CV < 1),
                           R := "Stepper Motor ทำงาน สั่งconveyor เคลื่อที่ไปข้างหน้า" OR "ปุ่มClear",
                           PV := 1);
   IF "IEC_Counter_0_DB_875".Q THEN #Output := 395; END_IF;
   "IEC_Counter_0_DB_874".CTU(CU := ("ยา 396" = 1) AND ("IEC_Counter_0_DB_874".CV < 1),
                           R := "Stepper Motor ทำงาน สั่งconveyor เคลื่อที่ไปข้างหน้า" OR "ปุ่มClear",
                           PV := 1);
   IF "IEC_Counter_0_DB_874".Q THEN #Output := 396; END_IF;
   "IEC_Counter_0_DB_873".CTU(CU := ("ยา 397" = 1) AND ("IEC_Counter_0_DB_873".CV < 1),
                           R := "Stepper Motor ทำงาน สั่งconveyor เคลื่อที่ไปข้างหน้า" OR "ปุ่มClear",
                           PV := 1);
   IF "IEC_Counter_0_DB_873".Q THEN #Output := 397; END_IF;
   "IEC_Counter_0_DB_872".CTU(CU := ("ยา 398" = 1) AND ("IEC_Counter_0_DB_872".CV < 1),
                           R := "Stepper Motor ทำงาน สั่งconveyor เคลื่อที่ไปข้างหน้า" OR "ปุ่มClear",
                           PV := 1);
   IF "IEC_Counter_0_DB_872".Q THEN #Output := 398; END_IF;
   "IEC_Counter_0_DB_871".CTU(CU := ("ยา 399" = 1) AND ("IEC_Counter_0_DB_871".CV < 1),
                           R := "Stepper Motor ทำงาน สั่งconveyor เคลื่อที่ไปข้างหน้า" OR "ปุ่มClear",
                           PV := 1);
   IF "IEC_Counter_0_DB_871".Q THEN #Output := 399; END_IF;
   "IEC_Counter_0_DB_870".CTU(CU := ("ยา 400" = 1) AND ("IEC_Counter_0_DB_870".CV < 1),
                           R := "Stepper Motor ทำงาน สั่งconveyor เคลื่อที่ไปข้างหน้า" OR "ปุ่มClear",
                           PV := 1);
   IF "IEC_Counter_0_DB_870".Q THEN #Output := 400; END_IF;
END_REGION

REGION Network 21
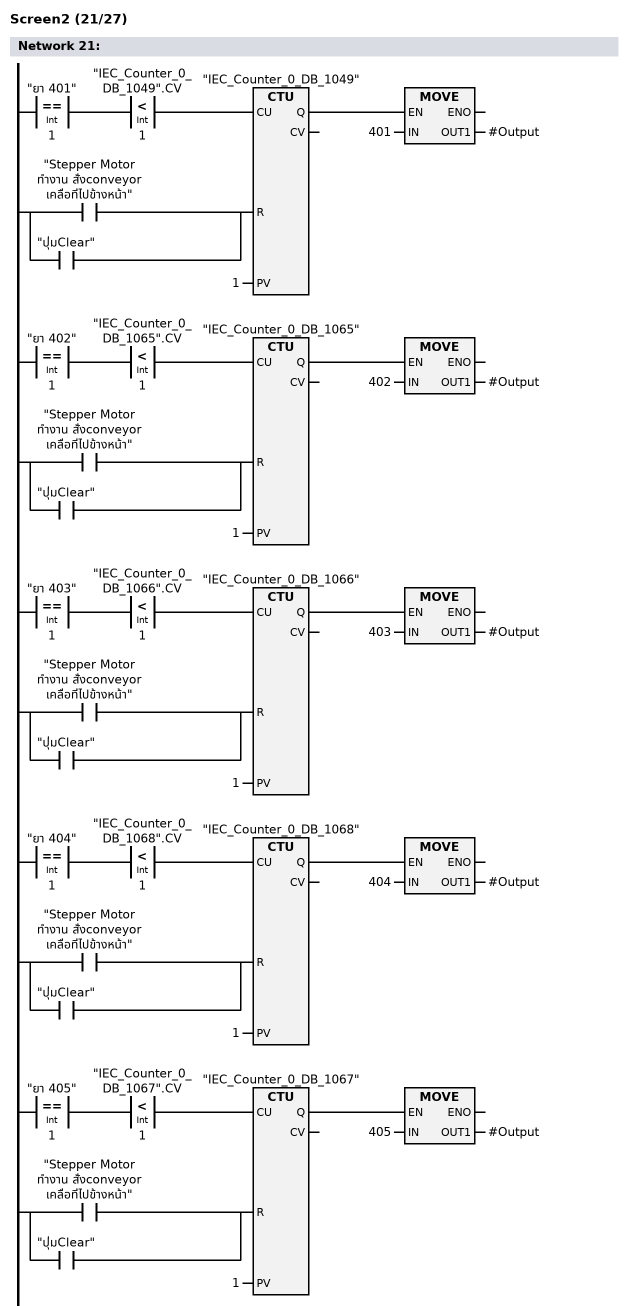
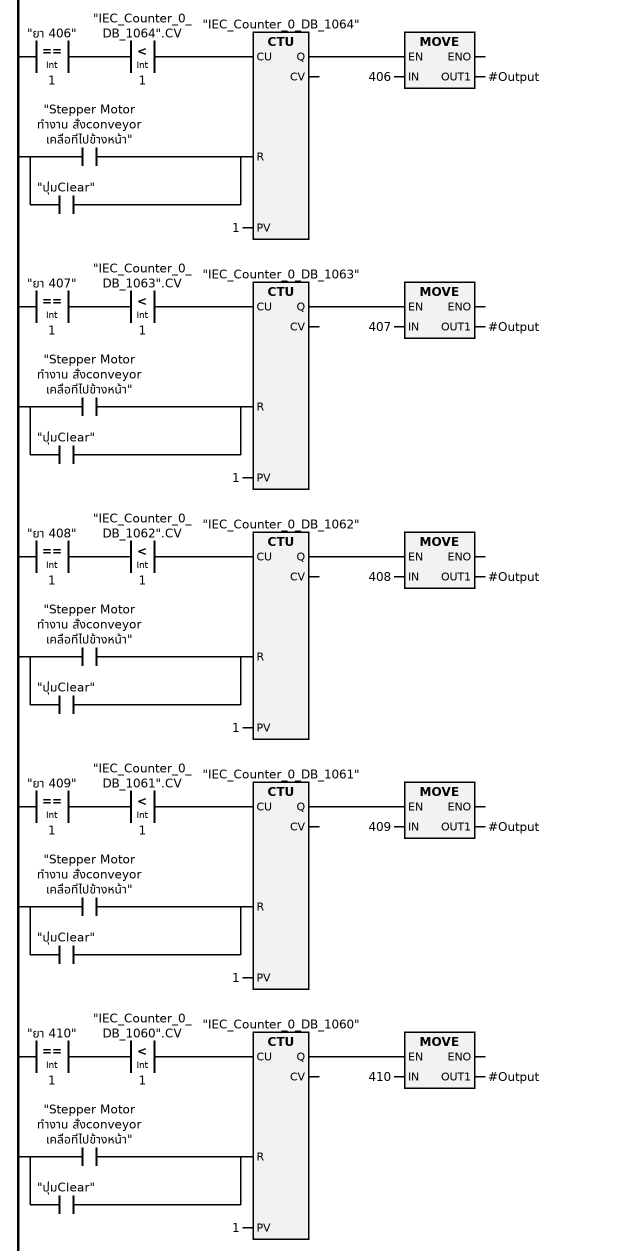
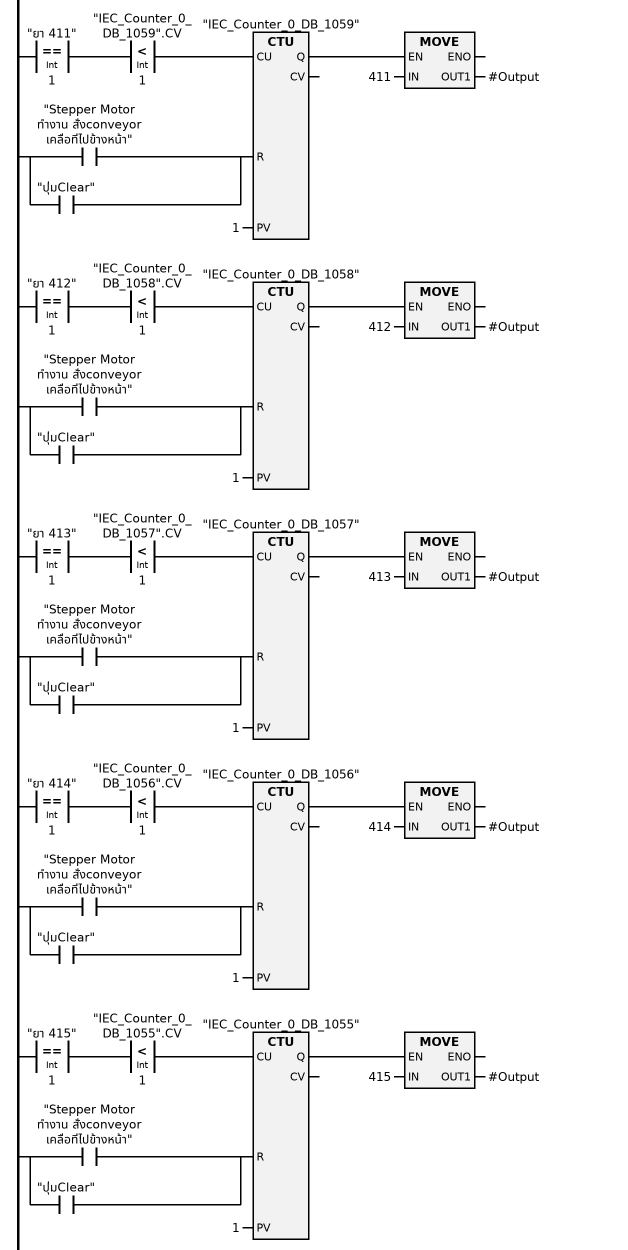
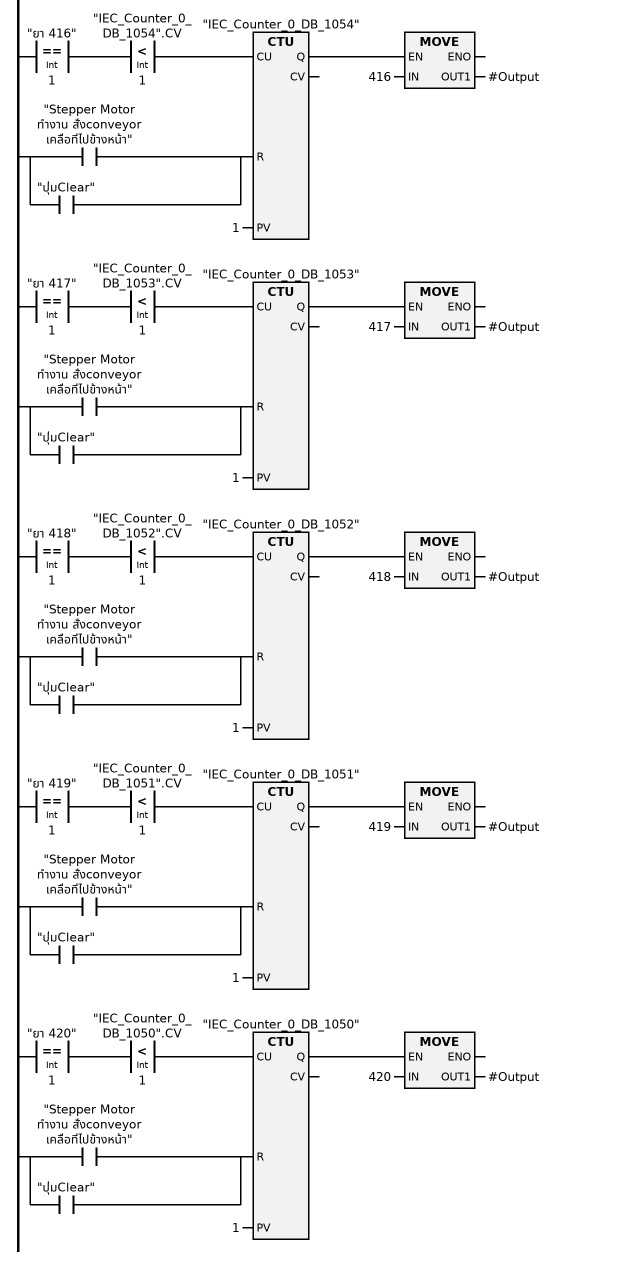
   "IEC_Counter_0_DB_1049".CTU(CU := ("ยา 401" = 1) AND ("IEC_Counter_0_DB_1049".CV < 1),
                           R := "Stepper Motor ทำงาน สั่งconveyor เคลื่อที่ไปข้างหน้า" OR "ปุ่มClear",
                           PV := 1);
   IF "IEC_Counter_0_DB_1049".Q THEN #Output := 401; END_IF;
   "IEC_Counter_0_DB_1065".CTU(CU := ("ยา 402" = 1) AND ("IEC_Counter_0_DB_1065".CV < 1),
                           R := "Stepper Motor ทำงาน สั่งconveyor เคลื่อที่ไปข้างหน้า" OR "ปุ่มClear",
                           PV := 1);
   IF "IEC_Counter_0_DB_1065".Q THEN #Output := 402; END_IF;
   "IEC_Counter_0_DB_1066".CTU(CU := ("ยา 403" = 1) AND ("IEC_Counter_0_DB_1066".CV < 1),
                           R := "Stepper Motor ทำงาน สั่งconveyor เคลื่อที่ไปข้างหน้า" OR "ปุ่มClear",
                           PV := 1);
   IF "IEC_Counter_0_DB_1066".Q THEN #Output := 403; END_IF;
   "IEC_Counter_0_DB_1068".CTU(CU := ("ยา 404" = 1) AND ("IEC_Counter_0_DB_1068".CV < 1),
                           R := "Stepper Motor ทำงาน สั่งconveyor เคลื่อที่ไปข้างหน้า" OR "ปุ่มClear",
                           PV := 1);
   IF "IEC_Counter_0_DB_1068".Q THEN #Output := 404; END_IF;
   "IEC_Counter_0_DB_1067".CTU(CU := ("ยา 405" = 1) AND ("IEC_Counter_0_DB_1067".CV < 1),
                           R := "Stepper Motor ทำงาน สั่งconveyor เคลื่อที่ไปข้างหน้า" OR "ปุ่มClear",
                           PV := 1);
   IF "IEC_Counter_0_DB_1067".Q THEN #Output := 405; END_IF;
   "IEC_Counter_0_DB_1064".CTU(CU := ("ยา 406" = 1) AND ("IEC_Counter_0_DB_1064".CV < 1),
                           R := "Stepper Motor ทำงาน สั่งconveyor เคลื่อที่ไปข้างหน้า" OR "ปุ่มClear",
                           PV := 1);
   IF "IEC_Counter_0_DB_1064".Q THEN #Output := 406; END_IF;
   "IEC_Counter_0_DB_1063".CTU(CU := ("ยา 407" = 1) AND ("IEC_Counter_0_DB_1063".CV < 1),
                           R := "Stepper Motor ทำงาน สั่งconveyor เคลื่อที่ไปข้างหน้า" OR "ปุ่มClear",
                           PV := 1);
   IF "IEC_Counter_0_DB_1063".Q THEN #Output := 407; END_IF;
   "IEC_Counter_0_DB_1062".CTU(CU := ("ยา 408" = 1) AND ("IEC_Counter_0_DB_1062".CV < 1),
                           R := "Stepper Motor ทำงาน สั่งconveyor เคลื่อที่ไปข้างหน้า" OR "ปุ่มClear",
                           PV := 1);
   IF "IEC_Counter_0_DB_1062".Q THEN #Output := 408; END_IF;
   "IEC_Counter_0_DB_1061".CTU(CU := ("ยา 409" = 1) AND ("IEC_Counter_0_DB_1061".CV < 1),
                           R := "Stepper Motor ทำงาน สั่งconveyor เคลื่อที่ไปข้างหน้า" OR "ปุ่มClear",
                           PV := 1);
   IF "IEC_Counter_0_DB_1061".Q THEN #Output := 409; END_IF;
   "IEC_Counter_0_DB_1060".CTU(CU := ("ยา 410" = 1) AND ("IEC_Counter_0_DB_1060".CV < 1),
                           R := "Stepper Motor ทำงาน สั่งconveyor เคลื่อที่ไปข้างหน้า" OR "ปุ่มClear",
                           PV := 1);
   IF "IEC_Counter_0_DB_1060".Q THEN #Output := 410; END_IF;
   "IEC_Counter_0_DB_1059".CTU(CU := ("ยา 411" = 1) AND ("IEC_Counter_0_DB_1059".CV < 1),
                           R := "Stepper Motor ทำงาน สั่งconveyor เคลื่อที่ไปข้างหน้า" OR "ปุ่มClear",
                           PV := 1);
   IF "IEC_Counter_0_DB_1059".Q THEN #Output := 411; END_IF;
   "IEC_Counter_0_DB_1058".CTU(CU := ("ยา 412" = 1) AND ("IEC_Counter_0_DB_1058".CV < 1),
                           R := "Stepper Motor ทำงาน สั่งconveyor เคลื่อที่ไปข้างหน้า" OR "ปุ่มClear",
                           PV := 1);
   IF "IEC_Counter_0_DB_1058".Q THEN #Output := 412; END_IF;
   "IEC_Counter_0_DB_1057".CTU(CU := ("ยา 413" = 1) AND ("IEC_Counter_0_DB_1057".CV < 1),
                           R := "Stepper Motor ทำงาน สั่งconveyor เคลื่อที่ไปข้างหน้า" OR "ปุ่มClear",
                           PV := 1);
   IF "IEC_Counter_0_DB_1057".Q THEN #Output := 413; END_IF;
   "IEC_Counter_0_DB_1056".CTU(CU := ("ยา 414" = 1) AND ("IEC_Counter_0_DB_1056".CV < 1),
                           R := "Stepper Motor ทำงาน สั่งconveyor เคลื่อที่ไปข้างหน้า" OR "ปุ่มClear",
                           PV := 1);
   IF "IEC_Counter_0_DB_1056".Q THEN #Output := 414; END_IF;
   "IEC_Counter_0_DB_1055".CTU(CU := ("ยา 415" = 1) AND ("IEC_Counter_0_DB_1055".CV < 1),
                           R := "Stepper Motor ทำงาน สั่งconveyor เคลื่อที่ไปข้างหน้า" OR "ปุ่มClear",
                           PV := 1);
   IF "IEC_Counter_0_DB_1055".Q THEN #Output := 415; END_IF;
   "IEC_Counter_0_DB_1054".CTU(CU := ("ยา 416" = 1) AND ("IEC_Counter_0_DB_1054".CV < 1),
                           R := "Stepper Motor ทำงาน สั่งconveyor เคลื่อที่ไปข้างหน้า" OR "ปุ่มClear",
                           PV := 1);
   IF "IEC_Counter_0_DB_1054".Q THEN #Output := 416; END_IF;
   "IEC_Counter_0_DB_1053".CTU(CU := ("ยา 417" = 1) AND ("IEC_Counter_0_DB_1053".CV < 1),
                           R := "Stepper Motor ทำงาน สั่งconveyor เคลื่อที่ไปข้างหน้า" OR "ปุ่มClear",
                           PV := 1);
   IF "IEC_Counter_0_DB_1053".Q THEN #Output := 417; END_IF;
   "IEC_Counter_0_DB_1052".CTU(CU := ("ยา 418" = 1) AND ("IEC_Counter_0_DB_1052".CV < 1),
                           R := "Stepper Motor ทำงาน สั่งconveyor เคลื่อที่ไปข้างหน้า" OR "ปุ่มClear",
                           PV := 1);
   IF "IEC_Counter_0_DB_1052".Q THEN #Output := 418; END_IF;
   "IEC_Counter_0_DB_1051".CTU(CU := ("ยา 419" = 1) AND ("IEC_Counter_0_DB_1051".CV < 1),
                           R := "Stepper Motor ทำงาน สั่งconveyor เคลื่อที่ไปข้างหน้า" OR "ปุ่มClear",
                           PV := 1);
   IF "IEC_Counter_0_DB_1051".Q THEN #Output := 419; END_IF;
   "IEC_Counter_0_DB_1050".CTU(CU := ("ยา 420" = 1) AND ("IEC_Counter_0_DB_1050".CV < 1),
                           R := "Stepper Motor ทำงาน สั่งconveyor เคลื่อที่ไปข้างหน้า" OR "ปุ่มClear",
                           PV := 1);
   IF "IEC_Counter_0_DB_1050".Q THEN #Output := 420; END_IF;
END_REGION

REGION Network 22
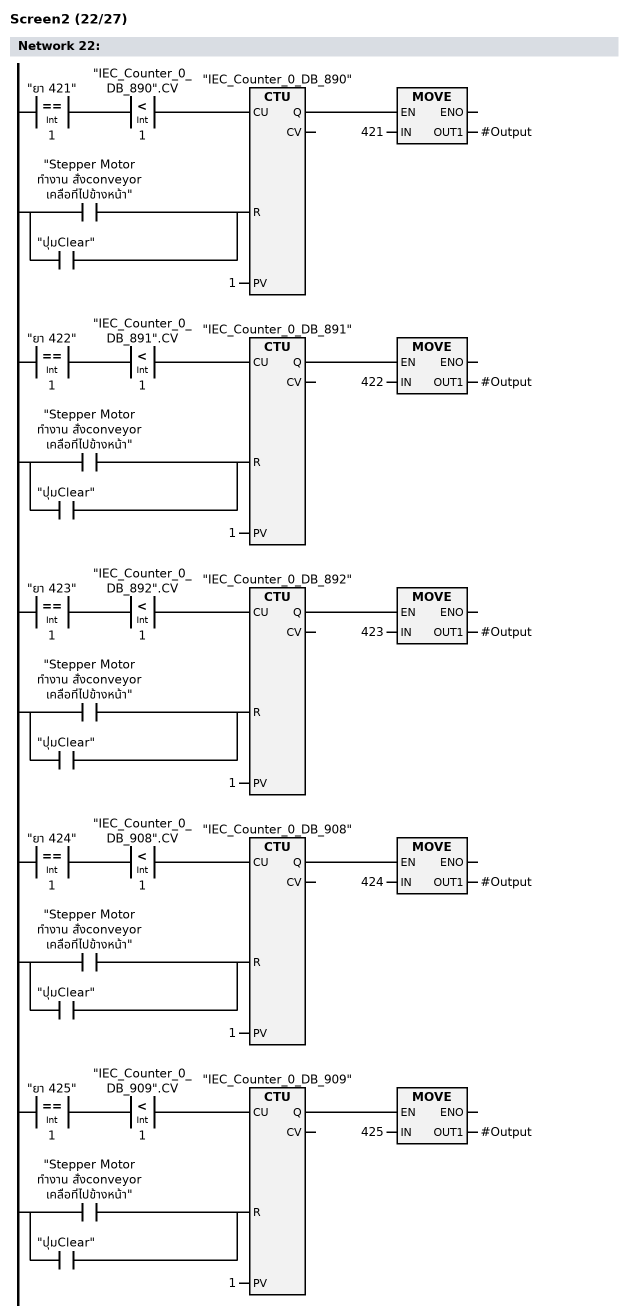
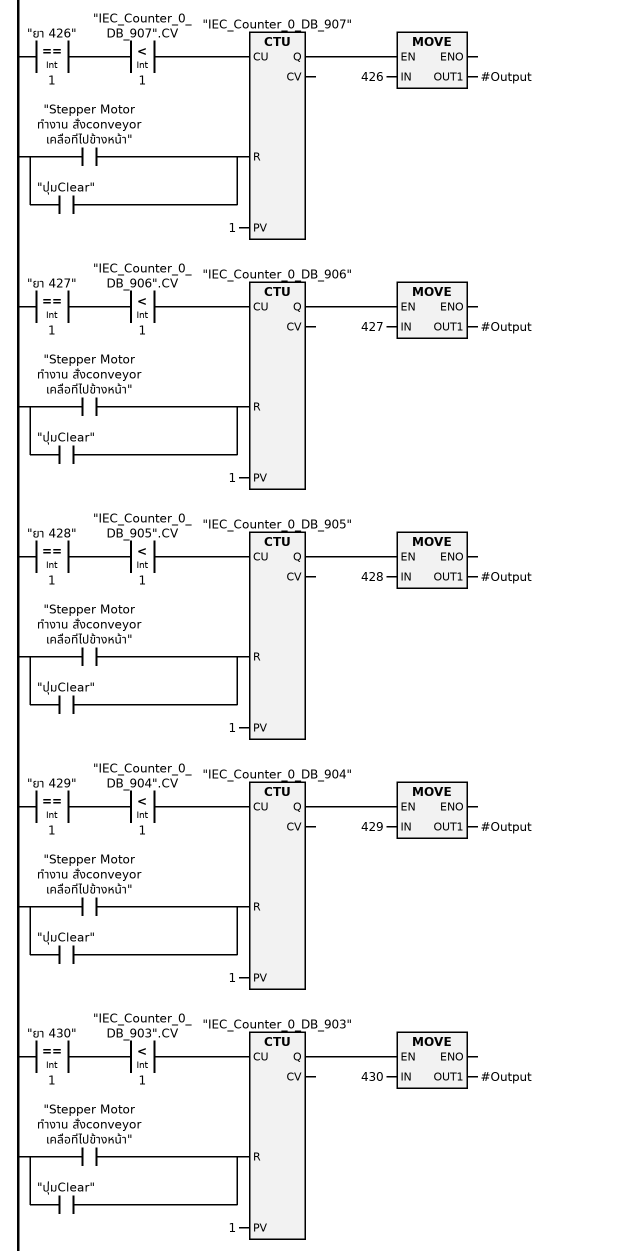
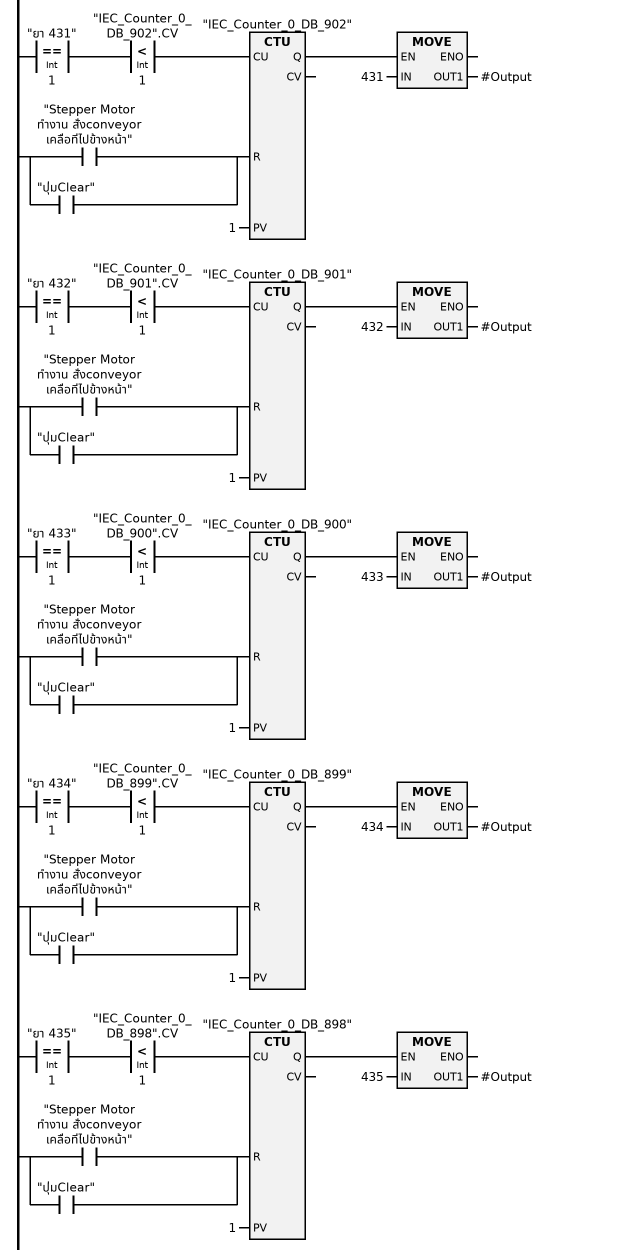
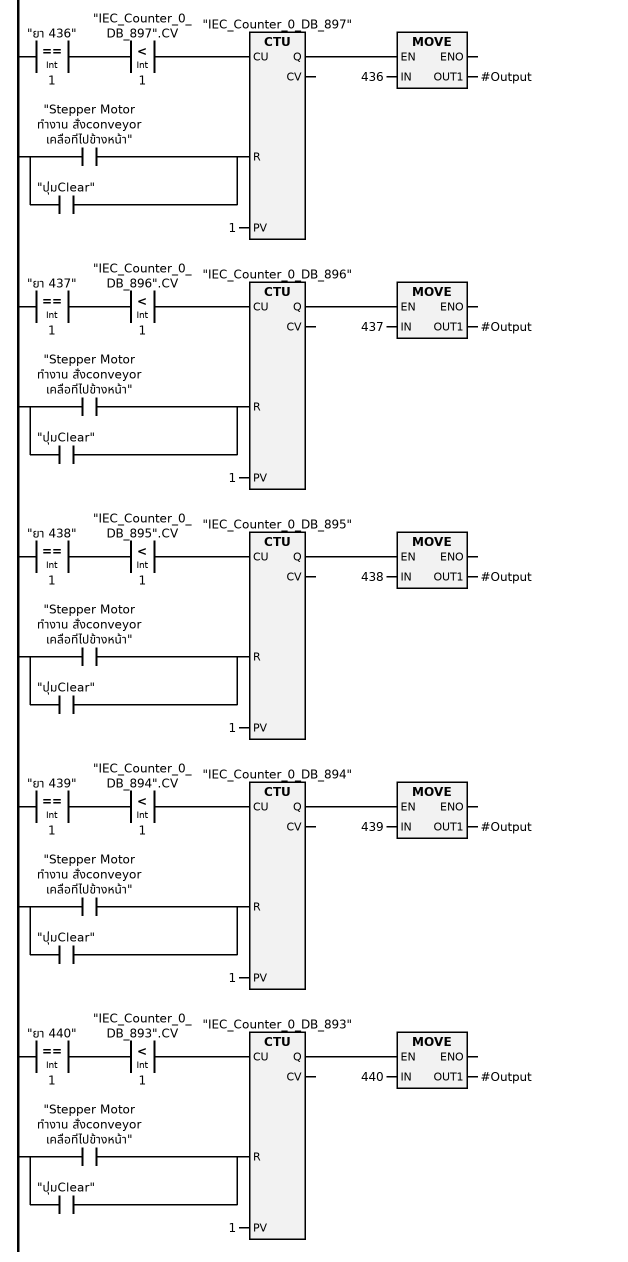
   "IEC_Counter_0_DB_890".CTU(CU := ("ยา 421" = 1) AND ("IEC_Counter_0_DB_890".CV < 1),
                           R := "Stepper Motor ทำงาน สั่งconveyor เคลื่อที่ไปข้างหน้า" OR "ปุ่มClear",
                           PV := 1);
   IF "IEC_Counter_0_DB_890".Q THEN #Output := 421; END_IF;
   "IEC_Counter_0_DB_891".CTU(CU := ("ยา 422" = 1) AND ("IEC_Counter_0_DB_891".CV < 1),
                           R := "Stepper Motor ทำงาน สั่งconveyor เคลื่อที่ไปข้างหน้า" OR "ปุ่มClear",
                           PV := 1);
   IF "IEC_Counter_0_DB_891".Q THEN #Output := 422; END_IF;
   "IEC_Counter_0_DB_892".CTU(CU := ("ยา 423" = 1) AND ("IEC_Counter_0_DB_892".CV < 1),
                           R := "Stepper Motor ทำงาน สั่งconveyor เคลื่อที่ไปข้างหน้า" OR "ปุ่มClear",
                           PV := 1);
   IF "IEC_Counter_0_DB_892".Q THEN #Output := 423; END_IF;
   "IEC_Counter_0_DB_908".CTU(CU := ("ยา 424" = 1) AND ("IEC_Counter_0_DB_908".CV < 1),
                           R := "Stepper Motor ทำงาน สั่งconveyor เคลื่อที่ไปข้างหน้า" OR "ปุ่มClear",
                           PV := 1);
   IF "IEC_Counter_0_DB_908".Q THEN #Output := 424; END_IF;
   "IEC_Counter_0_DB_909".CTU(CU := ("ยา 425" = 1) AND ("IEC_Counter_0_DB_909".CV < 1),
                           R := "Stepper Motor ทำงาน สั่งconveyor เคลื่อที่ไปข้างหน้า" OR "ปุ่มClear",
                           PV := 1);
   IF "IEC_Counter_0_DB_909".Q THEN #Output := 425; END_IF;
   "IEC_Counter_0_DB_907".CTU(CU := ("ยา 426" = 1) AND ("IEC_Counter_0_DB_907".CV < 1),
                           R := "Stepper Motor ทำงาน สั่งconveyor เคลื่อที่ไปข้างหน้า" OR "ปุ่มClear",
                           PV := 1);
   IF "IEC_Counter_0_DB_907".Q THEN #Output := 426; END_IF;
   "IEC_Counter_0_DB_906".CTU(CU := ("ยา 427" = 1) AND ("IEC_Counter_0_DB_906".CV < 1),
                           R := "Stepper Motor ทำงาน สั่งconveyor เคลื่อที่ไปข้างหน้า" OR "ปุ่มClear",
                           PV := 1);
   IF "IEC_Counter_0_DB_906".Q THEN #Output := 427; END_IF;
   "IEC_Counter_0_DB_905".CTU(CU := ("ยา 428" = 1) AND ("IEC_Counter_0_DB_905".CV < 1),
                           R := "Stepper Motor ทำงาน สั่งconveyor เคลื่อที่ไปข้างหน้า" OR "ปุ่มClear",
                           PV := 1);
   IF "IEC_Counter_0_DB_905".Q THEN #Output := 428; END_IF;
   "IEC_Counter_0_DB_904".CTU(CU := ("ยา 429" = 1) AND ("IEC_Counter_0_DB_904".CV < 1),
                           R := "Stepper Motor ทำงาน สั่งconveyor เคลื่อที่ไปข้างหน้า" OR "ปุ่มClear",
                           PV := 1);
   IF "IEC_Counter_0_DB_904".Q THEN #Output := 429; END_IF;
   "IEC_Counter_0_DB_903".CTU(CU := ("ยา 430" = 1) AND ("IEC_Counter_0_DB_903".CV < 1),
                           R := "Stepper Motor ทำงาน สั่งconveyor เคลื่อที่ไปข้างหน้า" OR "ปุ่มClear",
                           PV := 1);
   IF "IEC_Counter_0_DB_903".Q THEN #Output := 430; END_IF;
   "IEC_Counter_0_DB_902".CTU(CU := ("ยา 431" = 1) AND ("IEC_Counter_0_DB_902".CV < 1),
                           R := "Stepper Motor ทำงาน สั่งconveyor เคลื่อที่ไปข้างหน้า" OR "ปุ่มClear",
                           PV := 1);
   IF "IEC_Counter_0_DB_902".Q THEN #Output := 431; END_IF;
   "IEC_Counter_0_DB_901".CTU(CU := ("ยา 432" = 1) AND ("IEC_Counter_0_DB_901".CV < 1),
                           R := "Stepper Motor ทำงาน สั่งconveyor เคลื่อที่ไปข้างหน้า" OR "ปุ่มClear",
                           PV := 1);
   IF "IEC_Counter_0_DB_901".Q THEN #Output := 432; END_IF;
   "IEC_Counter_0_DB_900".CTU(CU := ("ยา 433" = 1) AND ("IEC_Counter_0_DB_900".CV < 1),
                           R := "Stepper Motor ทำงาน สั่งconveyor เคลื่อที่ไปข้างหน้า" OR "ปุ่มClear",
                           PV := 1);
   IF "IEC_Counter_0_DB_900".Q THEN #Output := 433; END_IF;
   "IEC_Counter_0_DB_899".CTU(CU := ("ยา 434" = 1) AND ("IEC_Counter_0_DB_899".CV < 1),
                           R := "Stepper Motor ทำงาน สั่งconveyor เคลื่อที่ไปข้างหน้า" OR "ปุ่มClear",
                           PV := 1);
   IF "IEC_Counter_0_DB_899".Q THEN #Output := 434; END_IF;
   "IEC_Counter_0_DB_898".CTU(CU := ("ยา 435" = 1) AND ("IEC_Counter_0_DB_898".CV < 1),
                           R := "Stepper Motor ทำงาน สั่งconveyor เคลื่อที่ไปข้างหน้า" OR "ปุ่มClear",
                           PV := 1);
   IF "IEC_Counter_0_DB_898".Q THEN #Output := 435; END_IF;
   "IEC_Counter_0_DB_897".CTU(CU := ("ยา 436" = 1) AND ("IEC_Counter_0_DB_897".CV < 1),
                           R := "Stepper Motor ทำงาน สั่งconveyor เคลื่อที่ไปข้างหน้า" OR "ปุ่มClear",
                           PV := 1);
   IF "IEC_Counter_0_DB_897".Q THEN #Output := 436; END_IF;
   "IEC_Counter_0_DB_896".CTU(CU := ("ยา 437" = 1) AND ("IEC_Counter_0_DB_896".CV < 1),
                           R := "Stepper Motor ทำงาน สั่งconveyor เคลื่อที่ไปข้างหน้า" OR "ปุ่มClear",
                           PV := 1);
   IF "IEC_Counter_0_DB_896".Q THEN #Output := 437; END_IF;
   "IEC_Counter_0_DB_895".CTU(CU := ("ยา 438" = 1) AND ("IEC_Counter_0_DB_895".CV < 1),
                           R := "Stepper Motor ทำงาน สั่งconveyor เคลื่อที่ไปข้างหน้า" OR "ปุ่มClear",
                           PV := 1);
   IF "IEC_Counter_0_DB_895".Q THEN #Output := 438; END_IF;
   "IEC_Counter_0_DB_894".CTU(CU := ("ยา 439" = 1) AND ("IEC_Counter_0_DB_894".CV < 1),
                           R := "Stepper Motor ทำงาน สั่งconveyor เคลื่อที่ไปข้างหน้า" OR "ปุ่มClear",
                           PV := 1);
   IF "IEC_Counter_0_DB_894".Q THEN #Output := 439; END_IF;
   "IEC_Counter_0_DB_893".CTU(CU := ("ยา 440" = 1) AND ("IEC_Counter_0_DB_893".CV < 1),
                           R := "Stepper Motor ทำงาน สั่งconveyor เคลื่อที่ไปข้างหน้า" OR "ปุ่มClear",
                           PV := 1);
   IF "IEC_Counter_0_DB_893".Q THEN #Output := 440; END_IF;
END_REGION

REGION Network 23
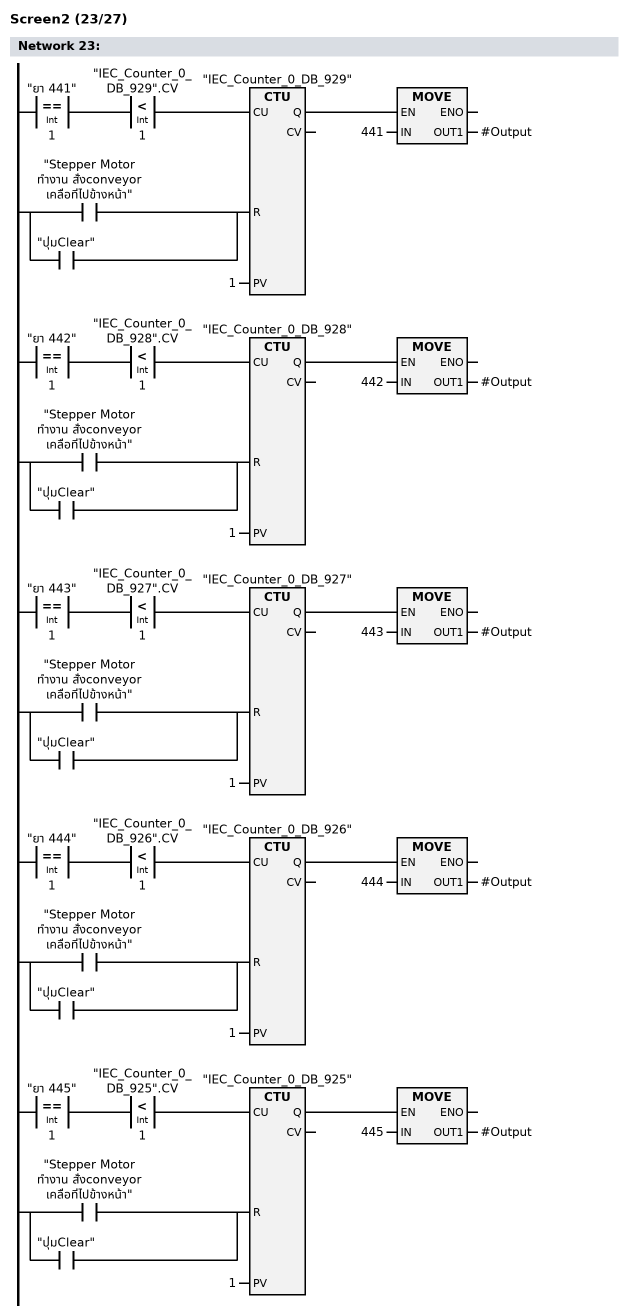
